(* IEC 61131-3 sources: daoli-st-library/DL_Process (part 20) *)

(* ---- FB_DL_AirShowerInterlockSeq.st ---- *)
(*
  ==================================================================
  组件名 Component  : FB_DL_AirShowerInterlockSeq
  分类   Category   : DL_Process
  复杂度 Complexity  : cx4
  版本   Version    : 1.0.0
  功能   Purpose    : 风淋室联锁顺控。双门互锁不变量（内 / 外门不得同时开，破坏
                      即故障锁存）；进入序列：外门开 → 外门关 → 吹淋计时 → 内门
                      许可 → 内门通过后回空闲；吹淋超时与中止（急停 / 火警电平）
                      优先解除全部门锁许可撤离；锁反馈校验失配判 eSensorBad。
  来源   Source     : t2-2-lbp（洁净室物流联锁族）
  溯源   Origin     : IEC 61131-3 标准语义的道莅防御性实现；双侧门 + 吹淋定时
                      三段联锁为通用洁净室语义，clean-room 自研实现，未复制任何
                      闭源代码行。
  平台   Platform   : 纯 IEC 61131-3（TON / R_TRIG / LREAL，无私有库）
  作者   Author     : 道莅代码库 · PLC 编程专家（R56）
  ------------------------------------------------------------------
  同拍双窗配比约束（R100）：tBlow（吹淋工艺窗）与 tBlowMax（吹淋看门狗窗）同相
                      并跑，配比约束 tBlowMax > tBlow 在组态域闸内判故障；
                      tFbTo 锁反馈失配消抖窗独立（不同相）。
  边界 Boundary     :
                      一 本件只出门锁与吹淋许可，不驱动门体电机、不控风机本体
                         （属主边界）；
                      二 安全侧优先：急停 / 火警电平（bEmgLevel）在任何相位立即
                         解除全部门锁并撤吹淋（撤离许可，安全侧直通）；
                      三 互锁不变量：bOuterLocked 与 bInnerLocked 不同拍同为假
                         （恒有一侧锁闭，双开即故障锁存）；
                      四 相级看门狗使能只用相驻留本身（R145）；
                      五 故障锁存解除路径 = bReset 上升沿（唯一路径，R188）；
                      六 无全局变量、无外部变量声明、无物理地址寻址。
  输出契约 Output contract:
                      bOuterLocked / bInnerLocked 为门锁命令电平（真 = 锁闭）；
                      bBlowing 为吹淋命令电平；bEntryAllowed 为进入许可（外门侧）；
                      eFault 为锁存回放；ePhaseBad 为非法相位兜底专用成员（R128）。
  修订记录 Revision  :
    2026-11-20  v1.0.0  R56 首版（批 4 · 序号 20）
  ==================================================================
*)

TYPE E_DL_AisPhase :
(
    eIdle       := 0,  // 空闲：外门侧许可进入 / idle, the outer side is allowed to enter
    eOuterOpen  := 10, // 外门开：人已进入，等外门关 / the outer door is open, waiting for it to close
    eBlow       := 20, // 吹淋：吹淋计时中，双侧门锁闭 / blowing, both doors locked
    eInnerAllow := 30, // 内门许可：吹淋完成，等内门通过 / the inner side allowed, waiting for the passage
    eAborted    := 40, // 已中止：全部门锁解除（撤离许可），等复位 / aborted, every lock released for evacuation
    eFault      := 90  // 故障：成因锁存，双侧解锁（安全侧）/ fault, the cause is latched with both sides unlocked
);
END_TYPE

TYPE E_DL_AisFault :
(
    eNone        := 0, // 无成因 / no cause
    eDoorBothOpen:= 1, // 双门同时开，互锁不变量被破坏（故障级，与 bError 配对）/ both doors open at once, the interlock invariant broken, fault grade paired with bError
    eBlowTimeout := 2, // 吹淋看门狗超时（故障级，与 bError 配对）/ the blow watchdog timed out, fault grade paired with bError
    eAborted     := 3, // 急停 / 火警中止（故障级，与 bError 配对）/ aborted by an emergency or fire level, fault grade paired with bError
    eSensorBad   := 4, // 锁反馈失配或组态非法（故障级，与 bError 配对）/ the lock feedback mismatches or the config illegal, fault grade paired with bError
    ePhaseBad    := 5  // 非法相位兜底（故障级，与 bError 配对）/ illegal phase fallback, fault grade paired with bError
);
END_TYPE

FUNCTION_BLOCK FB_DL_AirShowerInterlockSeq
VAR_INPUT
    bEnable      : BOOL := TRUE;    // 使能，失能时停顺控回空闲（门锁维持安全侧）[-] / enable, the sequence stops when disabled
    bReset       : BOOL := FALSE;   // 复位上升沿清故障锁存回空闲 [-] / reset rising edge clears the latch back to idle
    bOuterOpen   : BOOL := FALSE;   // 外门开反馈（真 = 开）[-] / the outer door open feedback, true is open
    bInnerOpen   : BOOL := FALSE;   // 内门开反馈（真 = 开）[-] / the inner door open feedback, true is open
    bOuterLockFb : BOOL := TRUE;    // 外门锁闭反馈（真 = 已锁）[-] / the outer lock feedback, true is locked
    bInnerLockFb : BOOL := TRUE;    // 内门锁闭反馈（真 = 已锁）[-] / the inner lock feedback, true is locked
    bEmgLevel    : BOOL := FALSE;   // 急停 / 火警电平（任何相位优先解除全部许可）[-] / the emergency or fire level, the top priority release
    tBlow        : TIME := T#15S;   // 吹淋工艺窗 [毫秒]，域 大于零 / the blow process window [millisecond], domain above zero
    tBlowMax     : TIME := T#30S;   // 吹淋看门狗窗 [毫秒]，域 大于 tBlow / the blow watchdog window, above the process window
    tPassTo      : TIME := T#30S;   // 内门通过超时窗 [毫秒]，域 大于零 / the inner passage timeout [millisecond], domain above zero
    tFbTo        : TIME := T#1S;    // 锁反馈失配消抖窗 [毫秒]，域 大于零 / the lock feedback mismatch debounce [millisecond], domain above zero
END_VAR
VAR_OUTPUT
    bOuterLocked  : BOOL := TRUE;  // 外门锁命令（真 = 锁闭）[-] / the outer lock command, true is locked
    bInnerLocked  : BOOL := TRUE;  // 内门锁命令（真 = 锁闭）[-] / the inner lock command, true is locked
    bBlowing      : BOOL := FALSE; // 吹淋命令电平 [-] / the blowing command level
    bEntryAllowed : BOOL := FALSE; // 进入许可（外门侧解锁派生）[-] / the entry permission, derived from the outer unlock
    ePhase        : E_DL_AisPhase := E_DL_AisPhase.eIdle; // 相位出口 [枚举] / phase outlet [enum]
    eFault        : E_DL_AisFault := E_DL_AisFault.eNone; // 成因出口，锁存回放 [枚举] / cause outlet replayed from the latch [enum]
    bError        : BOOL := FALSE; // 故障锁存标志 [-] / fault latch flag
END_VAR
VAR
    rtReset  : R_TRIG; // 复位沿检测，段 0 无条件刷新 / reset edge, refreshed unconditionally in segment zero
    tonBlow  : TON;    // 吹淋工艺窗，段 0 无条件刷新 / the blow process window, refreshed unconditionally
    tonBlowM : TON;    // 吹淋看门狗窗，段 0 无条件刷新 / the blow watchdog window, refreshed unconditionally
    tonPass  : TON;    // 内门通过超时窗，段 0 无条件刷新 / the inner passage timeout, refreshed unconditionally
    tonFb    : TON;    // 锁反馈失配消抖窗，段 0 无条件刷新 / the lock feedback mismatch debounce, refreshed unconditionally
    _ePhase  : E_DL_AisPhase := E_DL_AisPhase.eIdle; // 内部相位，CASE 唯一写入目标 / internal phase, the only CASE write target
    _eFaulC  : E_DL_AisFault := E_DL_AisFault.eNone; // 故障级成因，锁存至复位沿 / fault cause, latched until the reset edge
    _bFault  : BOOL := FALSE; // 故障锁存位 [-] / fault latch bit
    _bInit   : BOOL := FALSE; // 首扫初始化完成标志（R310）/ first scan initialisation flag
    _bCfgOk  : BOOL := FALSE; // 组态参数域内 [-] / the configuration is inside the domain
    _bFbBad  : BOOL := FALSE; // 锁反馈失配原始判据 [-] / the raw lock feedback mismatch verdict
END_VAR

// 段 0｜定时器与沿检测无条件周期刷新（禁入分支），IN 只串相位闸与状态闸（FB50-1）/ segment 0, unconditional refresh, no instance call inside a branch
rtReset(CLK := bReset); // 复位沿无条件刷新 / unconditional refresh of the reset edge
tonBlow(IN := (_ePhase = E_DL_AisPhase.eBlow) AND (NOT _bFault), PT := tBlow); // 吹淋工艺窗 / the blow process window
tonBlowM(IN := (_ePhase = E_DL_AisPhase.eBlow) AND (NOT _bFault), PT := tBlowMax); // 吹淋看门狗窗（R100：tBlowMax > tBlow 组态闸证明）/ the blow watchdog with the proven pairing
tonPass(IN := (_ePhase = E_DL_AisPhase.eInnerAllow) AND (NOT _bFault), PT := tPassTo); // 内门通过超时窗 / the inner passage timeout
tonFb(IN := _bFbBad AND (NOT _bFault), PT := tFbTo); // 锁反馈失配消抖窗 / the mismatch debounce

// 段 1｜首扫初始化（R310）/ segment 1, first scan initialisation
IF NOT _bInit THEN // 首扫一拍 / the very first scan
    _bInit := TRUE; // 置首扫完成标志 / raise the first scan flag
    _ePhase := E_DL_AisPhase.eIdle; // 相位从空闲起步 / the phase starts from idle
    _eFaulC := E_DL_AisFault.eNone; // 故障级成因清零 / clear the fault cause
    _bFault := FALSE; // 故障锁存清零 / clear the fault latch
END_IF

// 段 2｜复位沿作用域：清锁存 / 迁相位（门锁命令随相位派生重映射，两项逐项声明）/ segment 2, reset edge scope declared item by item
IF rtReset.Q THEN // 复位沿 / the reset edge
    _bFault := FALSE; // 作用域一：清故障锁存 / scope one, clear the fault latch
    _eFaulC := E_DL_AisFault.eNone; // 作用域一：清故障级成因 / scope one, clear the fault cause
    _ePhase := E_DL_AisPhase.eIdle; // 作用域二：迁回空闲相（门锁命令随相重派生）/ scope two, migrate back to idle, the lock commands re-derive
END_IF

// 段 3｜组态域闸（R151 全覆盖，含 R100 配比）/ segment 3, the configuration gate with the window pairing
_bCfgOk := (tBlow > T#0S) AND (tBlowMax > tBlow) AND (tPassTo > T#0S) AND (tFbTo > T#0S); // 组态参数域判定（tBlowMax > tBlow 为双窗配比，R100）/ the configuration verdict with the pairing

// 段 4｜失配原始判据：锁命令与锁反馈不一致（消抖窗承载 eSensorBad 归因）/ segment 4, the raw mismatch verdict, the debounce carries the sensor cause
_bFbBad := (bOuterLocked <> bOuterLockFb) OR (bInnerLocked <> bInnerLockFb) OR (NOT _bCfgOk); // 命令与反馈失配或组态非法 / the command and the feedback disagree or the config is illegal

// 段 5｜双开不变量判据：任何相位破坏即故障锁存（安全侧双侧解锁）/ segment 5, the both open invariant, any violation latches a fault with both sides unlocked
IF bOuterOpen AND bInnerOpen AND (NOT _bFault) THEN // 双门同开且未锁存 / both doors open while unlatched
    _bFault := TRUE; // 置故障锁存 / raise the fault latch
    _eFaulC := E_DL_AisFault.eDoorBothOpen; // 故障级成因（R45 配对 bError）/ the fault cause paired with bError
    _ePhase := E_DL_AisPhase.eFault; // 迁故障相 / migrate to the fault phase
END_IF

// 段 6｜急停 / 火警优先解除（安全侧直通，R146 立即终止）/ segment 6, the emergency takes the top priority, the immediate safe side release
IF bEmgLevel AND (NOT _bFault) THEN // 急停电平且未锁存 / the emergency level while unlatched
    _bFault := TRUE; // 置故障锁存 / raise the fault latch
    _eFaulC := E_DL_AisFault.eAborted; // 故障级成因（R45 配对 bError）/ the fault cause paired with bError
    _ePhase := E_DL_AisPhase.eFault; // 迁故障相 / migrate to the fault phase
END_IF

// 段 7｜相位机：ENUM + CASE，含 ELSE 非法相位兜底（R128）/ segment 7, the phase machine with an ELSE fallback
CASE _ePhase OF
E_DL_AisPhase.eIdle: // 空闲相：外门侧许可进入（外门解锁，内门锁闭）/ the idle phase, the outer side is allowed
    IF bEnable AND (NOT _bFault) AND bOuterOpen THEN // 外门开，进入序列启动 / the outer door opens and the entry sequence starts
        _ePhase := E_DL_AisPhase.eOuterOpen; // 迁外门开相 / migrate to the outer open phase
    END_IF

E_DL_AisPhase.eOuterOpen: // 外门开相：人已进入，等外门关（退出条件 ≥2：外门关 / 中止 / 失能 / 双开，R98）/ the outer open phase with at least two exit conditions
    IF (NOT bEnable) OR bEmgLevel THEN // 失能或急停 / disabled or an emergency
        _ePhase := E_DL_AisPhase.eFault; // 迁故障相（急停归因已在段 6 锁存）/ migrate to the fault phase
    ELSIF (NOT bOuterOpen) THEN // 外门已关 / the outer door has closed
        _ePhase := E_DL_AisPhase.eBlow; // 迁吹淋相 / migrate to the blow phase
    END_IF

E_DL_AisPhase.eBlow: // 吹淋相：双侧门锁闭，吹淋计时 / the blow phase, both doors locked and the timing runs
    IF (NOT bEnable) OR bEmgLevel THEN // 失能或急停 / disabled or an emergency
        _ePhase := E_DL_AisPhase.eFault; // 迁故障相 / migrate to the fault phase
    ELSIF tonBlowM.Q THEN // 看门狗超时（R100 看门狗窗）/ the watchdog expired
        _bFault := TRUE; // 置故障锁存 / raise the fault latch
        _eFaulC := E_DL_AisFault.eBlowTimeout; // 故障级成因（R45 配对 bError）/ the fault cause paired with bError
        _ePhase := E_DL_AisPhase.eFault; // 迁故障相 / migrate to the fault phase
    ELSIF tonBlow.Q THEN // 吹淋工艺窗完成（R80 三段：拍 N 进入序列起点 / 本拍行为：许可翻转 / 拍 N+1 转出：内门许可相）/ the process window completed
        _ePhase := E_DL_AisPhase.eInnerAllow; // 迁内门许可相 / migrate to the inner allow phase
    END_IF

E_DL_AisPhase.eInnerAllow: // 内门许可相：等内门通过（退出条件 ≥2：通过 / 超时 / 中止 / 失能，R98）/ the inner allow phase with at least two exit conditions
    IF (NOT bEnable) OR bEmgLevel THEN // 失能或急停 / disabled or an emergency
        _ePhase := E_DL_AisPhase.eFault; // 迁故障相 / migrate to the fault phase
    ELSIF NOT bInnerOpen THEN // 内门已关（人已通过）/ the inner door has closed, the passage is complete
        _ePhase := E_DL_AisPhase.eIdle; // 回空闲相（本批次结束，等待下一进入）/ back to idle for the next entry
    ELSIF tonPass.Q THEN // 内门通过超时 / the passage timed out
        _bFault := TRUE; // 置故障锁存 / raise the fault latch
        _eFaulC := E_DL_AisFault.eBlowTimeout; // 故障级成因（通过超时归并吹淋超时子带，R190 同带子带留痕）/ the fault cause, the passage timeout rides the blow band
        _ePhase := E_DL_AisPhase.eFault; // 迁故障相 / migrate to the fault phase
    END_IF

E_DL_AisPhase.eAborted: // 已中止相：全部解锁撤离许可，等复位沿 / the aborted phase, every lock released until the reset edge
    IF NOT bEnable THEN // 失能 / disabled
        _ePhase := E_DL_AisPhase.eIdle; // 迁未使能相 / migrate to idle
    END_IF

E_DL_AisPhase.eFault: // 故障相：成因锁存，等复位沿 / the fault phase, the cause is latched until the reset edge
    IF NOT bEnable THEN // 失能 / disabled
        _ePhase := E_DL_AisPhase.eIdle; // 迁未使能相 / migrate to idle
    END_IF

ELSE // 非法相位兜底（R128）/ the illegal phase fallback
    _bFault := TRUE; // 置故障锁存 / raise the fault latch
    _eFaulC := E_DL_AisFault.ePhaseBad; // 故障级成因（R45 配对 bError）/ the fault cause paired with bError
    _ePhase := E_DL_AisPhase.eFault; // 迁故障相 / migrate to the fault phase
END_CASE

// 段 8｜门锁与吹淋出口派生（互锁不变量的结构性承载 + eAborted 成员可达性）/ segment 8, the lock and blow outlets, the structural carrier
IF (_ePhase = E_DL_AisPhase.eAborted) OR (_ePhase = E_DL_AisPhase.eFault) THEN // 中止或故障相：双侧解锁撤离许可（安全侧）/ the aborted or fault phase, both sides unlock for evacuation
    bOuterLocked := FALSE; // 外门解锁 / the outer side unlocks
    bInnerLocked := FALSE; // 内门解锁 / the inner side unlocks
    bBlowing := FALSE; // 吹淋撤 / the blowing withdraws
ELSIF _ePhase = E_DL_AisPhase.eIdle THEN // 空闲相：外门侧许可 / the idle phase, the outer permission
    bOuterLocked := FALSE; // 外门解锁（进入许可）/ the outer side unlocks for entry
    bInnerLocked := TRUE; // 内门锁闭 / the inner side locks
    bBlowing := FALSE; // 吹淋撤 / the blowing withdraws
ELSIF _ePhase = E_DL_AisPhase.eOuterOpen THEN // 外门开相：双侧锁闭（人已在腔内）/ the outer open phase, both sides lock
    bOuterLocked := TRUE; // 外门锁闭 / the outer side locks
    bInnerLocked := TRUE; // 内门锁闭 / the inner side locks
    bBlowing := FALSE; // 吹淋撤 / the blowing withdraws
ELSIF _ePhase = E_DL_AisPhase.eBlow THEN // 吹淋相：双侧锁闭 + 吹淋 / the blow phase, both sides lock and the blowing runs
    bOuterLocked := TRUE; // 外门锁闭 / the outer side locks
    bInnerLocked := TRUE; // 内门锁闭 / the inner side locks
    bBlowing := TRUE; // 吹淋命令 / the blowing command
ELSE // 内门许可相：内门侧解锁 / the inner allow phase, the inner permission
    bOuterLocked := TRUE; // 外门锁闭 / the outer side locks
    bInnerLocked := FALSE; // 内门解锁（通过许可）/ the inner side unlocks for the passage
    bBlowing := FALSE; // 吹淋撤 / the blowing withdraws
END_IF
bEntryAllowed := (NOT bOuterLocked) AND (NOT _bFault); // 进入许可派生（故障否决）/ the entry permission derived with the fault veto

// 段 9｜反馈失配判级与统一出口 / segment 9, the feedback mismatch grading and the unified outlet
IF (NOT _bFault) AND tonFb.Q THEN // 失配消抖窗到且未锁存 / the debounce elapsed while unlatched
    _bFault := TRUE; // 置故障锁存 / raise the fault latch
    _eFaulC := E_DL_AisFault.eSensorBad; // 故障级成因（R45 配对 bError）/ the fault cause paired with bError
    _ePhase := E_DL_AisPhase.eFault; // 迁故障相 / migrate to the fault phase
END_IF
IF _bFault THEN // 故障锁存优先 / the fault latch takes priority
    eFault := _eFaulC; // 故障级成因锁存回放（R152）/ the fault cause replayed from the latch
ELSE
    eFault := E_DL_AisFault.eNone; // 无锁存即无成因 / no latch, no cause
END_IF
ePhase := _ePhase; // 相位出口单点映射 / single point phase outlet mapping
bError := _bFault; // 故障标志与锁存位同源 / the fault flag shares the latch source
END_FUNCTION_BLOCK

(* ---- FB_DL_AlarmShelving.st ---- *)
(*==============================================================================
 * 组件名称 (Component)  : FB_DL_AlarmShelving
 * 溯源说明 (Provenance) : 道莅 clean-room 防御性实现（ISA-18.2 族深化）
 * 所属子库 (Sublibrary) : DL_Process / AlarmGovernance
 * 当前版本 (Version)    : 1.0.0
 * 兼容性   (Platform)   : CODESYS 3.5 / TwinCAT 3 / 汇川 InoProShop；
 *                         纯 IEC 61131-3（第 3 版），仅用标准库 TON / R_TRIG
 * 组件分类 (Category)   : 功能块（FUNCTION_BLOCK）· 报警搁置管理（ISA-18.2 搁置态）
 * 功能一句话 (Summary)  : 限时搁置告警，超时强制恢复，搁置台账计数，与报警管理件正交。
 * 边界与安全 (Boundary) : ①无告警时搁置指令拒绝（台账不增，置码 035D）；
 *                         ②超时强制恢复优先于新搁置指令（同拍仲裁）；
 *                         ③搁置 TON 与指令沿检测无条件周期刷新；
 *                         ④bOut=告警态 AND NOT 搁置态（对下游呈现口径）；
 *                         ⑤超时恢复 bTimeout 为单拍脉冲，下一拍自清。
 * 错误码    : 16#0005_035D 无效搁置指令（无告警时搁置被拒）——信息级（单拍）
 *             16#0005_035E 搁置超时强制恢复——信息级（单拍脉冲）
 * 码位总账  : 16#0005_035D 用 / 16#0005_035E 用
 * 修改记录  : v1.0.0 R26 初版
 *==============================================================================*)
FUNCTION_BLOCK FB_DL_AlarmShelving
VAR_INPUT
    bAlarmActive : BOOL; // 原始告警态输入 / Raw alarm active input
    bShelveCmd   : BOOL; // 搁置指令（上升沿生效）/ Shelve command (rising edge)
    tMaxShelve   : TIME; // 最大搁置时长 [ms] / Maximum shelve duration [ms]
    bRestoreCmd  : BOOL; // 恢复指令（上升沿生效）/ Restore command (rising edge)
END_VAR
VAR_OUTPUT
    bOut         : BOOL; // 对下游呈现的告警态（搁置时 FALSE）/ Alarm state presented downstream
    bShelved     : BOOL; // 当前搁置态 / Currently shelved
    bTimeout     : BOOL; // 超时强制恢复单拍脉冲 / Timeout forced-restore one-shot pulse
    uShelveCount : UDINT; // 搁置台账累计计数 / Shelve ledger total count
    eErr         : UDINT; // 本周期错误码，0=无错 / Error code this cycle, 0 = none
END_VAR
VAR
    tonShelve : TON;   // 搁置计时（无条件刷新）/ Shelve timer, unconditional refresh
    rShelve   : R_TRIG; // 搁置指令上升沿（无条件刷新）/ Shelve command edge
    rRestore  : R_TRIG; // 恢复指令上升沿（无条件刷新）/ Restore command edge
    bTimeoutPulse: BOOL; // 超时单拍内部（锁存后下拍清）/ Timeout one-shot internal
END_VAR

// ---------- 无条件周期刷新：沿检测与搁置计时 ----------
rShelve (CLK := bShelveCmd);
rRestore(CLK := bRestoreCmd);
tonShelve(IN := bShelved, PT := tMaxShelve);

// ---------- 周期起点：错误码与超时脉冲先清（单拍生命周期） ----------
eErr := 0;
bTimeout := FALSE;

// ---------- 超时强制恢复：优先于新搁置指令（同拍仲裁） ----------
IF tonShelve.Q THEN
    bShelved := FALSE;                        // 强制恢复 / Forced restore
    bTimeoutPulse := TRUE;                    // 超时脉冲锁存 / Timeout pulse latched
    uShelveCount := uShelveCount + UDINT#1;   // 台账记一次超时 / Ledger counts timeout
END_IF

// ---------- 搁置指令仲裁 ----------
IF rShelve.Q THEN
    IF bAlarmActive AND (NOT bShelved) THEN
        bShelved := TRUE;                     // 有效搁置 / Valid shelve
        uShelveCount := uShelveCount + UDINT#1; // 台账计数加一 / Ledger increment
    ELSE
        eErr := 16#0005_035D;                 // 无效搁置（无告警或已搁置）/ Invalid shelve
    END_IF
END_IF

// ---------- 恢复指令仲裁（人工恢复） ----------
IF rRestore.Q AND bShelved THEN
    bShelved := FALSE;                        // 人工恢复 / Manual restore
END_IF

// ---------- 超时单拍脉冲：置位后下一拍清零（先出后清） ----------
IF bTimeoutPulse THEN
    bTimeout := TRUE;                            // 本拍输出超时脉冲 / Timeout pulse this cycle
    bTimeoutPulse := FALSE;                   // 内部单拍自销 / Internal one-shot self-clear
END_IF

// ---------- 对下游呈现口径：原始告警被搁置时呈现为无告警 ----------
bOut := bAlarmActive AND (NOT bShelved);

END_FUNCTION_BLOCK

(* ---- FB_DL_AmcMonitorStat.st ---- *)
(*
  ==================================================================
  组件名 Component  : FB_DL_AmcMonitorStat
  分类   Category   : DL_Process
  版本   Version    : 1.0.0
  功能   Purpose    : AMC 污染在线统计分级。在周期采样窗内累计气态分子污染浓度
                      （单位 ppb）的样本数、均值、峰值与超阈比例，窗末按三级阈
                      （A / B / C）把均值定级为 A / B / C / D 四档，C 档及以下
                      置报警；同时给出本窗超阈样本比例与连续超阈窗计数。
  溯源   Origin     : AMC 分级统计为洁净室污染监控的通用口径；本件为 clean-room
                      实现，仅借鉴来源分类与参数域组织（来源标签 roadmap-p2-amc），
                      道莅原创设计，未复制任何闭源代码行。
  平台   Platform   : 纯 IEC 61131-3（TON / REAL 运算，无私有库、无方言转换）
  作者   Author     : 道莅代码库 · PLC 编程专家（R55）
  ------------------------------------------------------------------
  边界 Boundary     :
                      一 本件只做统计分级与报警，不控制新风阀、不驱动净化设备（属主边界）；
                      二 采样窗由自复位周期 TON 驱动，窗末结算并清零累加器；
                      三 非有限浓度样本不参与统计，只累加坏样本计数（信息级，不置故障）；
                      四 三级阈必须严格递增，否则判组态故障并锁存至复位沿；
                      五 无全局变量、无外部变量声明、无物理地址寻址。
  输出契约 Output contract:
                      eClass 四档互斥，仅在窗末结算拍更新（锁存至下一窗末）；
                      bAlarm 在 C 档及以下（含 D 档）为真，挂状态量不挂单拍标志；
                      fMeanPpb / fMaxPpb / fExceedPct 为上一完整窗的结算值；
                      eCause 故障级成因与 bError 配对（R45），信息级永不置 bError。
  修订记录 Revision  :
    2026-11-20  v1.0.0  R55 首版（批 3 · 序号 13）
  ==================================================================
*)

TYPE E_DL_AmcClass :
(
    eA := 0,            // A 档：均值不高于 A 级阈 / class A, the mean stays at or below the A limit
    eB := 10,           // B 档：均值高于 A 级阈但不高于 B 级阈 / class B, above the A limit and at or below the B limit
    eC := 20,           // C 档：均值高于 B 级阈但不高于 C 级阈 / class C, above the B limit and at or below the C limit
    eD := 30            // D 档：均值高于 C 级阈 / class D, above the C limit
);
END_TYPE

TYPE E_DL_AmcCause :
(
    eNone       := 0,   // 无成因 / no cause
    eCfgIllegal := 1,   // 组态非法：三级阈非严格递增或比例阈越域（故障级，与 bError 配对）/ illegal config, limits not strictly increasing or the ratio threshold out of domain
    eBadSample  := 2,   // 存在非有限样本，未参与统计（信息级）/ non-finite samples excluded from the statistics, informational
    eNoSample   := 3    // 本窗无有效样本，等级保持上窗值（信息级）/ no valid sample in the window and the class holds, informational
);
END_TYPE

FUNCTION_BLOCK FB_DL_AmcMonitorStat
VAR_INPUT
    bEnable     : BOOL := TRUE;              // 使能，失能时冻结统计与等级 [-] / enable, the statistics and the class freeze when disabled
    bReset      : BOOL := FALSE;            // 复位上升沿清故障锁存与统计 [-] / reset rising edge clears the fault latch and the statistics
    fAmcPpb     : REAL := 0.0;               // AMC 浓度实测 [ppb] / measured AMC concentration [ppb]
    fClsALimit  : REAL := 10.0;              // A 级阈 [ppb]，域 大于零 / class A limit [ppb], domain above zero
    fClsBLimit  : REAL := 50.0;              // B 级阈 [ppb]，须大于 A 级阈 / class B limit [ppb], must exceed the class A limit
    fClsCLimit  : REAL := 100.0;             // C 级阈 [ppb]，须大于 B 级阈 / class C limit [ppb], must exceed the class B limit
    fExceedPctLimit : REAL := 20.0;          // 超阈样本比例报警阈 [百分比]，域 0..100 / exceed ratio alarm threshold [percent], domain 0 to 100
    tSampleWin  : TIME := T#60S;             // 采样窗时长 [毫秒]，域 大于零 / sampling window duration [millisecond], domain above zero
END_VAR
VAR_OUTPUT
    fMeanPpb    : REAL := 0.0;               // 上一窗均值 [ppb] / mean of the last complete window [ppb]
    fMaxPpb     : REAL := 0.0;               // 上一窗峰值 [ppb] / peak of the last complete window [ppb]
    fExceedPct  : REAL := 0.0;               // 上一窗超阈样本比例 [百分比] / exceed sample ratio of the last complete window [percent]
    nSampleCnt  : INT := 0;                  // 上一窗有效样本数 [个] / valid sample count of the last complete window
    nBadSampleCnt : INT := 0;                // 上一窗坏样本数 [个] / bad sample count of the last complete window
    nExceedWinCnt : INT := 0;                // 连续超比例窗计数（饱和到上限）[窗] / consecutive exceed windows, saturated [window]
    eClass      : E_DL_AmcClass := E_DL_AmcClass.eA; // 等级出口 [枚举] / class outlet [enum]
    bAlarm      : BOOL := FALSE;             // 报警（C 档及以下）[-] / alarm for class C and below
    bWinDone    : BOOL := FALSE;             // 窗结算单拍脉冲 [-] / window settle single-shot pulse
    eCause      : E_DL_AmcCause := E_DL_AmcCause.eNone; // 成因出口 [枚举] / cause outlet [enum]
    bError      : BOOL := FALSE;             // 故障锁存标志 [-] / fault latch flag
END_VAR
VAR
    rtReset     : R_TRIG;                    // 复位沿检测，段 0 无条件刷新 / reset edge detector, refreshed unconditionally in segment zero
    tonWin      : TON;                       // 采样窗周期计时（自复位式）/ sampling window timer, self resetting
    _eCause     : E_DL_AmcCause := E_DL_AmcCause.eNone;  // 信息级成因，每拍重算 / informational cause, recomputed every scan
    _eFaultCause: E_DL_AmcCause := E_DL_AmcCause.eNone;  // 故障级成因，锁存至复位沿 / fault cause, latched until the reset edge
    _eClass     : E_DL_AmcClass := E_DL_AmcClass.eA;     // 等级锁存量 / latched class
    _bFault     : BOOL := FALSE;             // 故障锁存位 [-] / fault latch bit
    _bInit      : BOOL := FALSE;             // 首扫初始化完成标志（R310）/ first scan initialisation flag
    _bSampleOk  : BOOL := FALSE;             // 本拍样本有限 [-] / this scan sample finite
    _bCfgBad    : BOOL := FALSE;             // 组态非法判定 [-] / illegal configuration verdict
    _bBadSeen   : BOOL := FALSE;             // 本窗出现过坏样本 [-] / a bad sample occurred in this window
    _bDoneInt   : BOOL := FALSE;             // 窗结算脉冲内部位，统一出口映射 / internal window done bit, mapped at the unified outlet
    _nCnt       : INT := 0;                  // 本窗有效样本计数 [个] / valid sample count of this window
    _nBad       : INT := 0;                  // 本窗坏样本计数 [个] / bad sample count of this window
    _nExceed    : INT := 0;                  // 本窗超阈样本计数 [个] / exceed sample count of this window
    _nExceedWin : INT := 0;                  // 连续超比例窗计数 [窗] / consecutive exceed window count [window]
    _nBadLast   : INT := 0;                  // 上一窗坏样本数锁存 [个] / last window bad sample count
    _nCntLast   : INT := 0;                  // 上一窗有效样本数锁存 [个] / last window valid sample count
    _fSum       : REAL := 0.0;               // 本窗浓度累加 [ppb] / concentration sum of this window [ppb]
    _fMax       : REAL := 0.0;               // 本窗浓度峰值 [ppb] / concentration peak of this window [ppb]
    _fMean      : REAL := 0.0;               // 本窗均值工作值 [ppb] / mean working value of this window [ppb]
    _fExceedPct : REAL := 0.0;               // 本窗超阈比例工作值 [百分比] / exceed ratio working value [percent]
    _fMeanLast  : REAL := 0.0;               // 上一窗均值锁存 [ppb] / last window mean
    _fMaxLast   : REAL := 0.0;               // 上一窗峰值锁存 [ppb] / last window peak
    _fExcLast   : REAL := 0.0;               // 上一窗超阈比例锁存 [百分比] / last window exceed ratio
END_VAR
VAR CONSTANT
    DL_AMC_WIN_MIN   : REAL := 0.0;          // 浓度下限（负浓度不可能）[ppb] / concentration floor, negatives are impossible [ppb]
    DL_AMC_WIN_MAX   : REAL := 1.0E6;        // 浓度量级上限，防量纲错配 [ppb] / concentration magnitude ceiling against a mismatch [ppb]
    DL_AMC_PCT_MAX   : REAL := 100.0;        // 比例上限 [百分比] / ratio ceiling [percent]
    DL_AMC_CNT_MAX   : INT := 30000;         // 单窗样本计数上限，防溢出 [个] / per window sample count ceiling against overflow [count]
    DL_AMC_WIN_CNT_MAX : INT := 10000;       // 连续超比例窗计数上限 [窗] / consecutive exceed window count ceiling [window]
END_VAR

// 段 0｜定时器与沿检测无条件周期刷新（禁入分支）；采样窗用自复位式（IN 取自身 Q 的补）/ segment 0, unconditional refresh with a self resetting window timer
rtReset(CLK := bReset); // 复位沿无条件刷新 / unconditional refresh of the reset edge
tonWin(IN := (NOT tonWin.Q) AND bEnable AND (NOT _bFault), PT := tSampleWin); // 周期窗自复位：Q 到时下一拍 IN 变假即重启，符合周期脉冲发生器用法（不得用于闭锁窗）/ self resetting periodic window, never used as a latching window

// 段 1｜首扫初始化（R310）/ segment 1, first scan initialisation
IF NOT _bInit THEN // 首扫一拍 / the very first scan
    _bInit := TRUE; // 置首扫完成标志 / raise the first scan flag
    _bFault := FALSE; // 故障锁存清零 / clear the fault latch
    _eCause := E_DL_AmcCause.eNone; // 信息级成因清零 / clear the informational cause
    _eFaultCause := E_DL_AmcCause.eNone; // 故障级成因清零 / clear the fault cause
    _eClass := E_DL_AmcClass.eA; // 等级从 A 档起步 / the class starts at A
    _nCnt := 0; // 有效样本计数清零 / clear the valid sample count
    _nBad := 0; // 坏样本计数清零 / clear the bad sample count
    _nExceed := 0; // 超阈计数清零 / clear the exceed count
    _fSum := 0.0; // 浓度累加清零 / clear the concentration sum
    _fMax := 0.0; // 峰值清零 / clear the peak
END_IF

// 段 2｜复位沿作用域：清锁存 / 清统计 / 清等级（三项逐项声明）/ segment 2, reset edge scope
IF rtReset.Q THEN // 复位沿 / reset edge
    _bFault := FALSE; // 作用域一：清故障锁存 / scope one, clear the fault latch
    _eFaultCause := E_DL_AmcCause.eNone; // 作用域一：清故障级成因 / scope one, clear the fault cause
    _nCnt := 0; // 作用域二：清有效样本计数 / scope two, clear the valid count
    _nBad := 0; // 作用域二：清坏样本计数 / scope two, clear the bad count
    _nExceed := 0; // 作用域二：清超阈计数 / scope two, clear the exceed count
    _fSum := 0.0; // 作用域二：清浓度累加 / scope two, clear the sum
    _fMax := 0.0; // 作用域二：清峰值 / scope two, clear the peak
    _nExceedWin := 0; // 作用域二：清连续超比例窗计数 / scope two, clear the consecutive exceed window count
    _eClass := E_DL_AmcClass.eA; // 作用域三：等级回 A 档 / scope three, the class returns to A
    _bDoneInt := FALSE; // 作用域一：清窗结算脉冲内部位 / scope one, clear the internal done bit
END_IF

// 段 3｜组态域闸（R151 全覆盖）：三级阈严格递增、比例阈域、窗时长 / segment 3, configuration domain gate with strictly increasing limits
_bCfgBad := FALSE; // 组态非法预置假 / preset the illegal configuration verdict to false
IF (fClsALimit <= DL_AMC_WIN_MIN) OR (fClsALimit <> fClsALimit) OR (fClsALimit > DL_AMC_WIN_MAX) THEN // A 级阈越域 / the A limit is out of domain
    _bCfgBad := TRUE; // 判非法 / mark illegal
END_IF
IF (fClsBLimit <= fClsALimit) OR (fClsBLimit <> fClsBLimit) OR (fClsBLimit > DL_AMC_WIN_MAX) THEN // B 级阈非大于 A 级阈 / the B limit is not above the A limit
    _bCfgBad := TRUE; // 判非法 / mark illegal
END_IF
IF (fClsCLimit <= fClsBLimit) OR (fClsCLimit <> fClsCLimit) OR (fClsCLimit > DL_AMC_WIN_MAX) THEN // C 级阈非大于 B 级阈 / the C limit is not above the B limit
    _bCfgBad := TRUE; // 判非法 / mark illegal
END_IF
IF (fExceedPctLimit < 0.0) OR (fExceedPctLimit > DL_AMC_PCT_MAX) OR (fExceedPctLimit <> fExceedPctLimit) THEN // 比例阈越域 / the ratio threshold is out of domain
    _bCfgBad := TRUE; // 判非法 / mark illegal
END_IF
IF tSampleWin <= T#0S THEN // 窗时长非正 / the window duration is not positive
    _bCfgBad := TRUE; // 判非法 / mark illegal
END_IF
IF _bCfgBad AND (NOT _bFault) THEN // 组态非法且未锁存 / illegal configuration and not yet latched
    _bFault := TRUE; // 置故障锁存 / raise the fault latch
    _eFaultCause := E_DL_AmcCause.eCfgIllegal; // 故障级成因 (R45 配对 bError) / fault grade cause paired with bError
END_IF

// 段 4｜样本接收：有限性与量级闸，坏样本不入统计 / segment 4, sample acceptance with finiteness and magnitude gates
_eCause := E_DL_AmcCause.eNone; // 信息级成因每拍重算 / the informational cause is recomputed every scan
_bSampleOk := (fAmcPpb = fAmcPpb) AND ((fAmcPpb - fAmcPpb) = (fAmcPpb - fAmcPpb)) AND (fAmcPpb >= DL_AMC_WIN_MIN) AND (fAmcPpb <= DL_AMC_WIN_MAX); // 样本有限性闸（NaN 自反、无穷差值自减）/ sample finiteness gate
IF bEnable AND (NOT _bFault) THEN // 使能且无故障才收样本 / samples are accepted only while enabled and unfaulted
    IF _bSampleOk THEN // 样本可用 / the sample is usable
        IF _nCnt < DL_AMC_CNT_MAX THEN // 未达计数上限 / below the count ceiling
            _nCnt := _nCnt + 1; // 有效样本计数递增 / increment the valid count
        END_IF
        _fSum := _fSum + fAmcPpb; // 浓度累加 / accumulate the concentration
        IF fAmcPpb > _fMax THEN // 峰值刷新 / refresh the peak
            _fMax := fAmcPpb; // 更新峰值 / update the peak
        END_IF
        IF fAmcPpb > fClsCLimit THEN // 超 C 级阈 / above the C limit
            IF _nExceed < DL_AMC_CNT_MAX THEN // 未达计数上限 / below the count ceiling
                _nExceed := _nExceed + 1; // 超阈计数递增 / increment the exceed count
            END_IF
        END_IF
    ELSE // 样本不可用 / the sample is unusable
        _bBadSeen := TRUE; // 记坏样本出现 / record the bad sample
        IF _nBad < DL_AMC_CNT_MAX THEN // 未达计数上限 / below the count ceiling
            _nBad := _nBad + 1; // 坏样本计数递增 / increment the bad count
        END_IF
    END_IF
END_IF

// 段 5｜窗末结算：算均值与超阈比例，定级并累加连续超比例窗 / segment 5, window settle with grading
IF tonWin.Q THEN // 窗末（自复位计时到时）/ window end
    _fMean := 0.0; // 均值预置零 / preset the mean to zero
    _fExceedPct := 0.0; // 超阈比例预置零 / preset the exceed ratio to zero
    IF _nCnt > 0 THEN // 有有效样本 / at least one valid sample
        _fMean := _fSum / INT_TO_REAL(_nCnt); // 均值，除子已证大于零 / mean, divisor proven positive
        _fExceedPct := INT_TO_REAL(_nExceed) / INT_TO_REAL(_nCnt) * 100.0; // 超阈比例，除子已证大于零 / exceed ratio, divisor proven positive
    END_IF
    _fMeanLast := _fMean; // 上一窗均值锁存 / latch the last window mean
    _fMaxLast := _fMax; // 上一窗峰值锁存 / latch the last window peak
    _fExcLast := _fExceedPct; // 上一窗比例锁存 / latch the last window ratio
    _nCntLast := _nCnt; // 上一窗样本数锁存 / latch the last window sample count
    _nBadLast := _nBad; // 上一窗坏样本数锁存 / latch the last window bad count
    IF _nCnt > 0 THEN // 有样本才定级 / grading needs samples
        IF _fMean <= fClsALimit THEN // 均值不高于 A 级阈 / the mean stays at or below the A limit
            _eClass := E_DL_AmcClass.eA; // A 档 / class A
        ELSIF _fMean <= fClsBLimit THEN // 高于 A 级阈且不高于 B 级阈 / above A and at or below B
            _eClass := E_DL_AmcClass.eB; // B 档 / class B
        ELSIF _fMean <= fClsCLimit THEN // 高于 B 级阈且不高于 C 级阈 / above B and at or below C
            _eClass := E_DL_AmcClass.eC; // C 档 / class C
        ELSE // 高于 C 级阈 / above the C limit
            _eClass := E_DL_AmcClass.eD; // D 档 / class D
        END_IF
        IF _fExceedPct > fExceedPctLimit THEN // 超阈比例超报警阈 / the exceed ratio passes the alarm threshold
            IF _nExceedWin < DL_AMC_WIN_CNT_MAX THEN // 未达计数上限 / below the ceiling
                _nExceedWin := _nExceedWin + 1; // 连续超比例窗计数递增 / increment the consecutive exceed window count
            END_IF
        ELSE
            _nExceedWin := 0; // 未超则清零 / cleared when the ratio is acceptable
        END_IF
    ELSE // 本窗无有效样本 / no valid sample this window
        _eCause := E_DL_AmcCause.eNoSample; // 信息级成因：等级保持上窗值 / informational cause, the class holds
    END_IF
    _bDoneInt := TRUE; // 窗结算脉冲内部位置位（统一出口映射，R187）/ raise the internal done bit, mapped at the unified outlet
    IF _bBadSeen THEN // 本窗出现过坏样本 / a bad sample occurred in this window
        _eCause := E_DL_AmcCause.eBadSample; // 信息级成因（坏样本比无样本更具体，后者不覆盖）/ informational cause, the bad sample is more specific than the empty window
    END_IF
    _bBadSeen := FALSE; // 坏样本标志按窗清零 / the bad sample flag is cleared per window
    // 累加器清零，进入下一窗 / clear the accumulators for the next window
    _nCnt := 0; // 有效样本计数清零 / clear the valid count
    _nBad := 0; // 坏样本计数清零 / clear the bad count
    _nExceed := 0; // 超阈计数清零 / clear the exceed count
    _fSum := 0.0; // 浓度累加清零 / clear the sum
    _fMax := 0.0; // 峰值清零 / clear the peak
END_IF
// 段 6｜统一出口 / segment 6, unified outlet
fMeanPpb := _fMeanLast; // 上一窗均值出口 / last window mean outlet
fMaxPpb := _fMaxLast; // 上一窗峰值出口 / last window peak outlet
fExceedPct := _fExcLast; // 上一窗比例出口 / last window ratio outlet
nSampleCnt := _nCntLast; // 上一窗样本数出口 / last window sample count outlet
nBadSampleCnt := _nBadLast; // 上一窗坏样本数出口 / last window bad count outlet
nExceedWinCnt := _nExceedWin; // 连续超比例窗计数出口 / consecutive exceed window count outlet
eClass := _eClass; // 等级出口（锁存量）/ class outlet from the latch
bAlarm := (_eClass = E_DL_AmcClass.eC) OR (_eClass = E_DL_AmcClass.eD); // 报警挂等级状态量（R99）/ the alarm follows the class state quantity
bWinDone := _bDoneInt; // 窗结算脉冲映射本拍值 / map the window done pulse for this scan
_bDoneInt := FALSE; // 映射后立即撤销，保证单拍宽度（R187 两段式）/ revoke right after mapping to keep a single-scan width
IF _bFault THEN // 故障锁存优先 / the fault latch takes priority
    eCause := _eFaultCause; // 故障级成因锁存回放 / the fault cause is replayed from the latch
ELSE
    eCause := _eCause; // 信息级成因直映 / the informational cause is mapped directly
END_IF
bError := _bFault; // 故障标志与锁存位同源 / the fault flag shares the latch source
END_FUNCTION_BLOCK

(* ---- FB_DL_AnaerobDigesterLoadCtrl.st ---- *)
(*
  道莅工业代码库 / Daoli Industrial ST Library
  组件: FB_DL_AnaerobDigesterLoadCtrl
  分类: DL_Process
  复杂度: C4 ｜ 版本: 1.0.0 ｜ 2026-11-24
  平台兼容: CODESYS 3.5+ / TwinCAT 3 / 汇川 InoProShop / 施耐德 Machine Expert
  开源溯源: 无（clean-room 工程算法自研；参考公开的厌氧消化 VFA/碱度比预警与产气量联动降载
            工艺经验，未复制任何受版权保护代码）
  许可证: 本项目自有 (MIT)

  功能职责:
    厌氧消化罐进料负荷控制。VFA/碱度比越限（>0.4）逐窗降载至下限 20% 流量；比值落回 0.25~0.4
    进 eWatch 保持不增；产气量低于基准 70% 连续确认后直接降载（码 41）；稳定后先一步 eDerate
    再进 eRecover，每窗回升 5% 直至回满并完成两级确认才回 eNormal。
    越限降载路径是安全侧：先降流量，再报码。

  输入/输出契约:
    IN  bEnable 上升沿启动（并做四项参数校验）；FALSE 输出归零回 eIdle（R191 声明）。
    IN  bReset 上升沿是 eFault 唯一出口（还须残留故障条件消失），同时流量归 0。
    OUT rFeedOutM3h 实际进料流量 = MIN(实测, 当前限值) [m3/h]。
    OUT iLoadLevel  0~10 级负荷显式映射（每 10% 限值一级），故障/空闲为 0 级。

  码表 (Codes):
    41 = 产气骤降联动降载（信息级；gas < 0.7×基准且基准有效）
    42 = 进料流量上限无效（故障级；rFeedMaxM3h ≤ 0 或非有限，限值与级数不可算）
    43 = 降载步长越域（信息级；rStepDownPct 越 (0,50] 已回默认 10%）
    44 = VFA/碱度比越限降载（信息级；ratio > 0.4）
    45 = 碱度无效（故障级；rAlkMgL ≤ 0，除零闸）
    46 = 关键入参非有限（故障级；vfa / gas / feed 任一 ABS > 1.0E15）
    47 = 产气基准未整定（信息级；产气联动降载已禁用，仅按比值控制，降级已声明）
    48 = 降至下限仍越限（故障级；已到 20% 流量下限而比值仍越限，需人工介入）
    99 = 非法状态枚举值（ELSE 兜底）

  边界与红线:
    ① 两个定时器与两个 R_TRIG 全在 CASE 外无条件刷新（R7），CASE 内只读 .Q。
    ② tonConfirm 覆盖 eNormal / eWatch / eDerate 三相（相位无关的越限累计窗），tonRecover 覆盖
       eDerate / eRecover 两相，二者均带 NOT .Q 自复位（R188），并在此显式声明为
       **跨相累计看门狗**（红线 14）——按相拆开会漏计跨相连续的越限/稳定，属判据缺陷。
    ③ 两级确认（防抖）：连续两个 tConfirm 窗都越限才降载（_iConfCnt 容量载体
       DL_ADC_CONF_MAX）；回升到 eNormal 亦须连续两个 tRecover 窗稳定且限值回满。
    ④ 降载步进单点执行（段 5 的 _bStepReq 触发器），每窗仅一步，禁在 CASE 分支内重复乘；
       降载下限 DL_ADC_FLOOR_RATIO = 20% 流量，上限回满 100%。
    ⑤ R528：bEnable 必须上升沿且碱度、流量上限、三项信号有效性都通过才迁 eNormal；
       全默认引脚时停留 eIdle，绝不直达 eNormal / eDerate。
    ⑥ eFault 出口 = rtReset.Q AND NOT _bFaultCondNow（逐码反算残留条件，R28 可达性）。
    ⑦ 派单原文「gas < 0.7*base 且 ABS(base)>FIN」中的 ABS(base)>FIN 若照写即为死谓词
       （基准不可能大于 1E15 才生效，等于永久禁用该降载路径）；此处按工程反证改写为
       「基准非零且有限」（_bBaseOk），并把「基准未整定」显式报码 47，不静默失效。
  修订历史: 2026-11-24  v1.0.0  R82-B 首版
*)

TYPE E_DL_AD_STATE :
(
    eIdle    := 0,    // 空闲：等使能上升沿 / Idle: waiting for the enable rising edge
    eNormal  := 1,    // 正常相：满负荷进料，持续监视 / Normal: full load feeding with continuous supervision
    eWatch   := 2,    // 关注相：比值 0.25~0.4，保持不增 / Watch: ratio between 0.25 and 0.4, hold and do not increase
    eDerate  := 3,    // 降载相：按窗步进降流量 / Derate: step the flow down window by window
    eRecover := 4,    // 回升相：每窗升 5% 直至回满 / Recover: raise five percent per window up to full load
    eFault   := 5     // 故障安全相：流量归零 / Fault safe phase: the flow is forced to zero
);
END_TYPE

FUNCTION_BLOCK FB_DL_AnaerobDigesterLoadCtrl
VAR_INPUT
    bEnable       : BOOL := FALSE;     // 使能（上升沿启动；FALSE 输出归零回空闲）/ Enable, rising edge starts, FALSE zeroes the outputs
    bReset        : BOOL := FALSE;     // 复位（上升沿，eFault 唯一出口，流量归零）/ Reset rising edge, the only fault exit, the flow is zeroed
    rVfaMgL       : REAL := 0.0;       // 挥发性脂肪酸 VFA [mg/L] / Volatile fatty acids [mg/L]
    rAlkMgL       : REAL := 0.0;       // 碱度（以 CaCO3 计）[mg/L] / Alkalinity as CaCO3 [mg/L]
    rGasM3h       : REAL := 0.0;       // 产气量实测 [m3/h] / Measured biogas flow [m3/h]
    rGasBaseM3h   : REAL := 0.0;       // 产气量基准（整定值）[m3/h] / Biogas flow baseline after commissioning [m3/h]
    rFeedM3h      : REAL := 0.0;       // 进料流量实测 [m3/h] / Measured feed flow [m3/h]
    rFeedMaxM3h   : REAL := 0.0;       // 进料流量上限（100% 负荷）[m3/h] / Feed flow upper limit at one hundred percent load [m3/h]
    rStepDownPct  : REAL := 10.0;      // 单次降载步长，有效域 (0,50] [%] / Per-step derate percentage, valid domain above zero up to fifty [%]
    tConfirm      : TIME := T#60S;     // 越限确认窗，有效域 1s..2h [s] / Violation confirmation window, valid domain 1s..2h [s]
    tRecover      : TIME := T#5M;      // 回升/稳定窗，有效域 1s..2h [s] / Recovery window, valid domain 1s..2h [s]
END_VAR
VAR_OUTPUT
    rFeedOutM3h   : REAL := 0.0;       // 实际进料流量设定 [m3/h] / Actual feed flow setpoint [m3/h]
    bFeedOn       : BOOL := FALSE;     // 进料运行位（故障相强制 FALSE）/ Feed run bit, forced FALSE in the fault phase
    iLoadLevel    : INT := 0;          // 负荷等级 0~10（每 10% 一级）[级] / Load level from zero to ten, one level per ten percent [level]
    iErrCode      : INT := 0;          // 错误码（故障期锁存回放）/ Error code, latched replay during fault
    sMsg          : STRING;            // 文本提示（当前相位摘要）/ Text message, a summary of the current phase
END_VAR
VAR
    _eState        : E_DL_AD_STATE := E_DL_AD_STATE.eIdle;   // 内部相位（CASE 唯一写入目标）/ Internal phase, the only CASE write target
    _bFaultLatch   : BOOL := FALSE;    // 故障锁存位 / Fault latch
    _iErrLatch     : INT := 0;         // 锁存故障码（故障期唯一回放源）/ Latched fault code, the only replay source during fault
    _iInfoCode     : INT := 0;         // 信息级码 / Info code
    _iErrTmp       : INT := 0;         // 当拍故障首因中间量 / First fault cause of this scan
    _bFaultReq     : BOOL := FALSE;    // 当拍故障请求（段 6 统一锁存）/ Fault request of this scan, latched at segment 6
    _bFaultCondNow : BOOL := FALSE;    // 残留故障条件（eFault 出口唯一附加判据）/ Residual fault condition, the only extra fault-exit criterion
    _bStepReq      : BOOL := FALSE;    // 本拍降载步请求（段 5 单点执行）/ Derate step request of this scan, executed once at segment 5
    _bStepOutDom   : BOOL := FALSE;    // 降载步长越域标志（本拍已回默认）/ Derate step out-of-domain flag, the default was applied this scan
    _bRatioOk      : BOOL := FALSE;    // 比值可算标志（碱度有效且有限）/ Ratio computable flag, alkalinity valid and finite
    _bBaseOk       : BOOL := FALSE;    // 产气基准有效标志（非零且有限）/ Biogas baseline valid flag, non-zero and finite
    _bViolation    : BOOL := FALSE;    // 越限标志（比值高 或 产气骤降）/ Violation flag, high ratio or a biogas collapse
    _bRatioHigh    : BOOL := FALSE;    // 比值越限标志（ratio > 0.4）/ High ratio flag
    _bRatioWatch   : BOOL := FALSE;    // 比值关注标志（0.25 < ratio ≤ 0.4）/ Watch band flag
    _bGasLow       : BOOL := FALSE;    // 产气骤降标志（gas < 0.7×基准）/ Biogas collapse flag
    _bStableCond   : BOOL := FALSE;    // 稳定条件（ratio < 0.25 且产气回 0.9×基准）/ Stable condition, low ratio and recovered gas
    _rVfaCl        : REAL := 0.0;      // VFA 净化副本 [mg/L] / Sanitised VFA copy [mg/L]
    _rAlkCl        : REAL := 0.0;      // 碱度净化副本 [mg/L] / Sanitised alkalinity copy [mg/L]
    _rGasCl        : REAL := 0.0;      // 产气净化副本 [m3/h] / Sanitised biogas copy [m3/h]
    _rFeedCl       : REAL := 0.0;      // 进料净化副本 [m3/h] / Sanitised feed copy [m3/h]
    _rFeedMax      : REAL := 0.0;      // 流量上限净化值 [m3/h] / Sanitised feed maximum [m3/h]
    _rRatio        : REAL := 0.0;      // VFA/碱度比（无量纲）/ VFA to alkalinity ratio, dimensionless
    _rStepPct      : REAL := 10.0;     // 生效降载步长 [%] / Effective derate step [%]
    _rStepRatio    : REAL := 0.1;      // 生效降载步长折比（无量纲）/ Effective derate step as a fraction, dimensionless
    _rFloorM3h     : REAL := 0.0;      // 流量下限 = 20% 上限 [m3/h] / Flow floor at twenty percent of the maximum [m3/h]
    _rFeedLimit    : REAL := 0.0;      // 当前流量限值 [m3/h] / Current feed flow limit [m3/h]
    _rLoadPct      : REAL := 0.0;      // 当前限值占上限百分比 [%] / Current limit as a percentage of the maximum [%]
    _iLevel        : INT := 0;         // 负荷等级中间量 [级] / Intermediate load level [level]
    _iConfCnt      : INT := 0;         // 连续越限窗计数，容量载体 DL_ADC_CONF_MAX [窗] / Consecutive violation windows, capacity carrier DL_ADC_CONF_MAX [window]
    _iRecovCnt     : INT := 0;         // 连续稳定窗计数，容量载体 DL_ADC_CONF_MAX [窗] / Consecutive stable windows, capacity carrier DL_ADC_CONF_MAX [window]
    _tConfirm      : TIME := T#60S;    // 越限确认窗钳定值 [s] / Clamped violation window [s]
    _tRecover      : TIME := T#5M;     // 回升窗钳定值 [s] / Clamped recovery window [s]
    rtReset        : R_TRIG;           // bReset 边沿（段 3 无条件刷新）/ bReset edge, refreshed unconditionally
    rtEnable       : R_TRIG;           // bEnable 边沿（段 3 无条件刷新，R528）/ bEnable edge, refreshed unconditionally
    tonConfirm     : TON;              // 越限累计窗（跨相看门狗，自复位）/ Cumulative violation window, cross-phase watchdog with self reset
    tonRecover     : TON;              // 稳定累计窗（跨相看门狗，自复位）/ Cumulative stable window, cross-phase watchdog with self reset
END_VAR
VAR CONSTANT
    DL_ADC_EPS         : REAL := 1.0E-6;   // 数值闸阈值 [-]/ Numeric guard threshold [-]
    DL_ADC_FIN         : REAL := 1.0E15;   // 非有限判据阈值（ABS 比较用）[-] / Non-finite criterion threshold, compared by ABS [-]
    DL_ADC_RATIO_HI    : REAL := 0.4;      // 比值越限阈值（无量纲）/ High ratio threshold, dimensionless
    DL_ADC_RATIO_LO    : REAL := 0.25;     // 比值正常阈值（无量纲）/ Low ratio threshold, dimensionless
    DL_ADC_GAS_DROP    : REAL := 0.7;      // 产气骤降判定比（无量纲）/ Biogas collapse factor, dimensionless
    DL_ADC_GAS_REC     : REAL := 0.9;      // 产气恢复判定比（无量纲）/ Biogas recovery factor, dimensionless
    DL_ADC_STEP_DEF    : REAL := 10.0;     // 降载步长默认值 [%] / Default derate step [%]
    DL_ADC_STEP_MAX    : REAL := 50.0;     // 降载步长上限 [%] / Derate step upper limit [%]
    DL_ADC_FLOOR_RATIO : REAL := 0.2;      // 流量下限折比 20%（无量纲）/ Flow floor fraction of twenty percent, dimensionless
    DL_ADC_STEP_UP     : REAL := 0.05;     // 回升每窗步长 5%（无量纲）/ Recovery step of five percent per window, dimensionless
    DL_ADC_PCT_BASE    : REAL := 100.0;    // 百分比基准 [%] / Percentage base [%]
    DL_ADC_CONF_MAX    : INT := 2;         // 两级确认所需连续窗数 [窗] / Consecutive windows needed for the two-stage confirmation [window]
    DL_ADC_LEVEL_MAX   : INT := 10;        // 负荷等级上限 [级] / Load level upper limit [level]
    DL_ADC_ONE         : INT := 1;         // 计数步进一 [1] / Counter step of one [1]
    DL_ADC_ZERO        : INT := 0;         // 计数零基准 [-] / Counter zero base [-]
    DL_ADC_T_MIN       : TIME := T#1S;     // 时间参数下限 [s] / Time parameter lower bound [s]
    DL_ADC_T_MAX       : TIME := T#2H;     // 时间参数上限 [s] / Time parameter upper bound [s]
    DL_ADC_T_CONF_DEF  : TIME := T#60S;    // 确认窗默认回退值（在域内）[s] / Default confirmation window inside the domain [s]
    DL_ADC_T_REC_DEF   : TIME := T#5M;     // 回升窗默认回退值（在域内）[s] / Default recovery window inside the domain [s]
END_VAR

(* —— 段 1：中间量预置（只清当拍扫描量，不清锁存/限值/窗计数，FB32-1） —— *)
_iErrTmp   := 0;                                     // 当拍故障首因复位 / Scan first fault cause reset
_bFaultReq := FALSE;                                 // 当拍故障请求复位 / Scan fault request reset
_bStepReq  := FALSE;                                 // 本拍降载步请求复位 / Derate step request reset

(* —— 段 2：时间参数两级回退 + 入参净化 + 判据量折算（组态域闸覆盖每个引脚） —— *)
IF (tConfirm < DL_ADC_T_MIN) OR (tConfirm > DL_ADC_T_MAX) THEN
    _tConfirm := DL_ADC_T_CONF_DEF;                  // 越域：回一级默认常量 / Out of domain: fall back to the default constant
ELSE
    _tConfirm := tConfirm;                           // 域内：原值采用 / Inside the domain: use as given
END_IF
IF (tRecover < DL_ADC_T_MIN) OR (tRecover > DL_ADC_T_MAX) THEN
    _tRecover := DL_ADC_T_REC_DEF;                   // 越域：回一级默认常量 / Out of domain: fall back to the default constant
ELSE
    _tRecover := tRecover;                           // 域内：原值采用 / Inside the domain: use as given
END_IF
_rVfaCl := rVfaMgL;                                  // VFA 净化副本 [mg/L] / Sanitised VFA copy [mg/L]
IF (ABS(_rVfaCl) > DL_ADC_FIN) OR (_rVfaCl < 0.0) THEN
    _rVfaCl := 0.0;                                  // 非有限或负值兜底为零 / Non-finite or negative falls back to zero
END_IF
_rAlkCl := rAlkMgL;                                  // 碱度净化副本 [mg/L] / Sanitised alkalinity copy [mg/L]
IF (ABS(_rAlkCl) > DL_ADC_FIN) OR (_rAlkCl < 0.0) THEN
    _rAlkCl := 0.0;                                  // 非有限或负值兜底为零 / Non-finite or negative falls back to zero
END_IF
_rGasCl := rGasM3h;                                  // 产气净化副本 [m3/h] / Sanitised biogas copy [m3/h]
IF (ABS(_rGasCl) > DL_ADC_FIN) OR (_rGasCl < 0.0) THEN
    _rGasCl := 0.0;                                  // 非有限或负值兜底为零 / Non-finite or negative falls back to zero
END_IF
_rFeedCl := rFeedM3h;                                // 进料净化副本 [m3/h] / Sanitised feed copy [m3/h]
IF (ABS(_rFeedCl) > DL_ADC_FIN) OR (_rFeedCl < 0.0) THEN
    _rFeedCl := 0.0;                                 // 非有限或负值兜底为零 / Non-finite or negative falls back to zero
END_IF
_rFeedMax := rFeedMaxM3h;                            // 流量上限净化值 [m3/h] / Sanitised feed maximum [m3/h]
IF (ABS(_rFeedMax) > DL_ADC_FIN) OR (_rFeedMax < 0.0) THEN
    _rFeedMax := 0.0;                                // 非有限或负值兜底为零 / Non-finite or negative falls back to zero
END_IF
_rStepPct := rStepDownPct;                           // 降载步长初值 [%] / Initial derate step [%]
_bStepOutDom := FALSE;                               // 越域标志预置 / Out-of-domain flag preset
IF (ABS(_rStepPct) > DL_ADC_FIN) OR (_rStepPct <= 0.0) OR (_rStepPct > DL_ADC_STEP_MAX) THEN
    _rStepPct    := DL_ADC_STEP_DEF;                 // 越域回默认（不静默：由信息码 43 上报）/ Out of domain falls back, reported by info code 43
    _bStepOutDom := TRUE;                            // 置越域标志（段 5 报码 43）/ Raise the flag, code 43 is emitted at segment 5
END_IF
_rStepRatio := _rStepPct / DL_ADC_PCT_BASE;          // 量纲: (%)/(%) = 无量纲折比 / Percentage over percentage gives a dimensionless fraction
_bRatioOk := (_rAlkCl > DL_ADC_EPS);                 // 比值可算：碱度有效（除零闸）/ The ratio is computable when the alkalinity is valid
IF _bRatioOk THEN
    // 量纲: (mg/L)/(mg/L) = 无量纲比值，与 0.4 / 0.25 无量纲阈值直比
    _rRatio := _rVfaCl / _rAlkCl;                    // VFA/碱度比（分母已闸）/ VFA to alkalinity ratio with a guarded denominator
ELSE
    _rRatio := 0.0;                                  // 分母无效：比值出零，绝不猜值 / Invalid denominator: the ratio is zero, never guessed
END_IF
_rFloorM3h := _rFeedMax * DL_ADC_FLOOR_RATIO;        // 量纲: (m3/h)*(无量纲) = m3/h 下限 / (m3/h) times dimensionless gives the floor [m3/h]
_bBaseOk := (ABS(rGasBaseM3h) > DL_ADC_EPS) AND (ABS(rGasBaseM3h) <= DL_ADC_FIN);   // 基准有效：非零且有限 / Baseline valid: non-zero and finite
_bRatioHigh  := _bRatioOk AND (_rRatio > DL_ADC_RATIO_HI);                                     // 比值越限 / High ratio
_bRatioWatch := _bRatioOk AND (_rRatio > DL_ADC_RATIO_LO) AND (NOT _bRatioHigh);                // 关注带 / Watch band
IF _bBaseOk THEN
    // 量纲: (m3/h)*(无量纲) = m3/h 判定门限
    _bGasLow     := _rGasCl < (rGasBaseM3h * DL_ADC_GAS_DROP);                                 // 产气骤降 / Biogas collapse
    _bStableCond := (_rRatio < DL_ADC_RATIO_LO) AND (_bRatioOk) AND (_rGasCl > (rGasBaseM3h * DL_ADC_GAS_REC));   // 稳定条件 / Stable condition
ELSE
    _bGasLow     := FALSE;                                                                      // 基准无效：产气联动禁用（码 47 上报）
    _bStableCond := (_rRatio < DL_ADC_RATIO_LO) AND (_bRatioOk);                                 // 仅按比值判定稳定 / Stability by ratio alone
END_IF
_bViolation := _bRatioHigh OR _bGasLow;              // 越限 = 比值高 或 产气骤降 / Violation is a high ratio or a biogas collapse
_bFaultCondNow := FALSE;                             // 残留条件预置（eFault 出口唯一附加判据）/ Residual preset, the only extra fault-exit criterion
IF _iErrLatch = 42 THEN
    _bFaultCondNow := (rFeedMaxM3h <= DL_ADC_EPS) OR (ABS(rFeedMaxM3h) > DL_ADC_FIN);   // 码 42：上限仍无效 / Code 42: the maximum is still invalid
ELSIF _iErrLatch = 45 THEN
    _bFaultCondNow := (rAlkMgL <= DL_ADC_EPS);                                          // 码 45：碱度仍无效 / Code 45: the alkalinity is still invalid
ELSIF _iErrLatch = 46 THEN
    _bFaultCondNow := (ABS(rVfaMgL) > DL_ADC_FIN) OR (ABS(rGasM3h) > DL_ADC_FIN) OR (ABS(rFeedM3h) > DL_ADC_FIN);   // 码 46：非有限仍在 / Code 46: the non-finite input persists
ELSIF _iErrLatch = 48 THEN
    _bFaultCondNow := _bViolation;                                                       // 码 48：越限仍在 / Code 48: the violation persists
END_IF
(* 码 99（非法枚举）为内部损坏，无输入残留条件，复位沿单独即可退出。 / Code 99 has no residual input condition *)

(* —— 段 3：边沿与定时器（全部在 CASE 外无条件刷新，R7；IN 带 NOT .Q 自复位，R188） —— *)
rtReset(CLK := bReset);                              // 复位边沿无条件刷新 / Reset edge refreshed unconditionally
rtEnable(CLK := bEnable);                            // 使能边沿无条件刷新（R528 起点判据）/ Enable edge refreshed unconditionally
tonConfirm(IN := ((_eState = E_DL_AD_STATE.eNormal) OR (_eState = E_DL_AD_STATE.eWatch)
                  OR (_eState = E_DL_AD_STATE.eDerate))
                 AND _bViolation AND (NOT tonConfirm.Q) AND (NOT _bFaultLatch),
           PT := _tConfirm);                         // 跨相累计看门狗：三相内越限持续累计，非本相超时 / Cumulative watchdog over three phases, not a phase timeout
tonRecover(IN := ((_eState = E_DL_AD_STATE.eDerate) OR (_eState = E_DL_AD_STATE.eRecover))
                 AND _bStableCond AND (NOT tonRecover.Q) AND (NOT _bFaultLatch),
           PT := _tRecover);                         // 跨相累计看门狗：降载与回升两相内稳定累计 / Cumulative watchdog over the derate and recover phases
IF NOT _bViolation THEN
    _iConfCnt := DL_ADC_ZERO;                        // 越限中断：连续窗计数清零（防抖前提）/ Violation interrupted: the consecutive window counter is cleared
END_IF
IF tonConfirm.Q THEN
    IF _iConfCnt < DL_ADC_CONF_MAX THEN
        _iConfCnt := _iConfCnt + DL_ADC_ONE;         // 越限窗计数 +1，达容量上限饱和 / Violation window counter incremented and saturated at capacity
    END_IF
END_IF
IF NOT _bStableCond THEN
    _iRecovCnt := DL_ADC_ZERO;                       // 稳定中断：连续窗计数清零 / Stability interrupted: the consecutive window counter is cleared
END_IF
IF tonRecover.Q THEN
    IF _iRecovCnt < DL_ADC_CONF_MAX THEN
        _iRecovCnt := _iRecovCnt + DL_ADC_ONE;       // 稳定窗计数 +1，达容量上限饱和 / Stable window counter incremented and saturated at capacity
    END_IF
END_IF

(* —— 段 4：状态机主体（唯一相位写入点；降载步只置请求，由段 5 单点执行） —— *)
CASE _eState OF
    E_DL_AD_STATE.eIdle :
        (* 迁移①：拍 N 进入（使能上升沿）/ 本拍行为：四项参数校验，缺任一即故障 / 拍 N+1 转出至正常相 *)
        IF rtEnable.Q AND (NOT _bFaultLatch) THEN
            IF (rFeedMaxM3h <= DL_ADC_EPS) OR (ABS(rFeedMaxM3h) > DL_ADC_FIN) THEN
                _iErrTmp   := 42;                                  // 故障级：流量上限无效 / Fault: invalid feed maximum
                _bFaultReq := TRUE;                                // 请求段 6 锁存 / Request the latch at segment 6
            ELSIF NOT _bRatioOk THEN
                _iErrTmp   := 45;                                  // 故障级：碱度无效（除零闸）/ Fault: invalid alkalinity
                _bFaultReq := TRUE;                                // 请求段 6 锁存 / Request the latch at segment 6
            ELSIF (ABS(rVfaMgL) > DL_ADC_FIN) OR (ABS(rGasM3h) > DL_ADC_FIN) OR (ABS(rFeedM3h) > DL_ADC_FIN) THEN
                _iErrTmp   := 46;                                  // 故障级：关键入参非有限 / Fault: a key input is non-finite
                _bFaultReq := TRUE;                                // 请求段 6 锁存 / Request the latch at segment 6
            ELSE
                _rFeedLimit := _rFeedMax;                          // 新周期：限值回满 100% / New cycle: the limit starts at one hundred percent
                _iConfCnt   := DL_ADC_ZERO;                        // 新周期：越限窗计数清零 / New cycle: violation window counter cleared
                _iRecovCnt  := DL_ADC_ZERO;                        // 新周期：稳定窗计数清零 / New cycle: stable window counter cleared
                _iInfoCode  := 0;                                  // 新周期：信息码归零 / New cycle: info code cleared
                IF NOT _bBaseOk THEN
                    _iInfoCode := 47;                              // 信息级：基准未整定，产气联动已禁用 / Info: no baseline, the biogas link is disabled
                END_IF
                _eState := E_DL_AD_STATE.eNormal;                  // 迁移①：进正常相 / Move to normal
            END_IF
        END_IF

    E_DL_AD_STATE.eNormal :
        (* 迁移②③④：拍 N 进入 / 本拍行为：满负荷监视；越限两级确认后降载 / 拍 N+1 转出 *)
        IF _iConfCnt >= DL_ADC_CONF_MAX THEN
            IF _bGasLow THEN
                _iInfoCode := 41;                                  // 信息级：产气骤降联动降载 / Info: biogas collapse derate
            ELSE
                _iInfoCode := 44;                                  // 信息级：比值越限降载 / Info: ratio violation derate
            END_IF
            _bStepReq := TRUE;                                     // 请求段 5 执行一步降载 / Request one derate step at segment 5
            _iRecovCnt := DL_ADC_ZERO;                             // 进降载：稳定窗计数清零 / Entering derate: the stable window counter is cleared
            _eState := E_DL_AD_STATE.eDerate;                      // 迁移②：进降载相 / Move to derate
        ELSIF _bRatioWatch THEN
            _iInfoCode := 0;                                       // 关注带不降载，仅保持不增 / The watch band does not derate, it only prevents increases
            _eState := E_DL_AD_STATE.eWatch;                        // 迁移③：进关注相 / Move to watch
        END_IF

    E_DL_AD_STATE.eWatch :
        (* 迁移⑤⑥：拍 N 进入 / 本拍行为：保持当前限值不增（禁回升）/ 拍 N+1 转出至降载相或正常相 *)
        IF _iConfCnt >= DL_ADC_CONF_MAX THEN
            IF _bGasLow THEN
                _iInfoCode := 41;                                  // 信息级：产气骤降联动降载 / Info: biogas collapse derate
            ELSE
                _iInfoCode := 44;                                  // 信息级：比值越限降载 / Info: ratio violation derate
            END_IF
            _bStepReq := TRUE;                                     // 请求段 5 执行一步降载 / Request one derate step at segment 5
            _iRecovCnt := DL_ADC_ZERO;                             // 进降载：稳定窗计数清零 / Entering derate: the stable window counter is cleared
            _eState := E_DL_AD_STATE.eDerate;                      // 迁移⑤：进降载相 / Move to derate
        ELSIF (_bRatioOk) AND (_rRatio < DL_ADC_RATIO_LO) THEN
            _eState := E_DL_AD_STATE.eNormal;                      // 迁移⑥：比值回落，回正常相 / Ratio recovered, back to normal
        END_IF

    E_DL_AD_STATE.eDerate :
        (* 迁移⑦⑧⑨：拍 N 进入 / 本拍行为：每个越限确认窗限速降一步 / 拍 N+1 转出至回升相或故障相 *)
        IF _rFeedLimit <= (_rFloorM3h + DL_ADC_EPS) THEN
            IF _bViolation THEN
                _iErrTmp   := 48;                                  // 故障级：已到下限仍越限 / Fault: still violating at the floor
                _bFaultReq := TRUE;                                // 请求段 6 锁存 / Request the latch at segment 6
            END_IF
        END_IF
        IF tonConfirm.Q AND (NOT _bFaultReq) THEN
            IF _bBaseOk AND _bGasLow THEN
                _iInfoCode := 41;                                  // 信息级：产气骤降继续降载 / Info: the biogas collapse keeps derating
            ELSIF _bRatioHigh THEN
                _iInfoCode := 44;                                  // 信息级：比值继续越限降载 / Info: the ratio keeps violating
            END_IF
            _bStepReq := TRUE;                                     // 请求段 5 再执行一步降载 / Request another derate step at segment 5
        END_IF
        IF tonRecover.Q THEN
            _eState := E_DL_AD_STATE.eRecover;                     // 迁移⑧：稳定一窗，进回升相 / One stable window, move to recover
        END_IF

    E_DL_AD_STATE.eRecover :
        (* 迁移⑩⑪⑫：拍 N 进入 / 本拍行为：每个稳定窗升 5%，回满且两级确认后回正常 / 拍 N+1 转出 *)
        IF _bViolation THEN
            _iConfCnt  := DL_ADC_ZERO;                             // 回升中越限：越限窗计数从头计 / Violation during recovery restarts the window counter
            _iInfoCode := 44;                                      // 信息级：回升中止（先降后报）/ Info: recovery aborted, derate first
            _bStepReq  := TRUE;                                    // 请求段 5 执行一步降载 / Request one derate step at segment 5
            _eState    := E_DL_AD_STATE.eDerate;                   // 迁移⑩：中止回升，回降载相 / Abort recovery and go back to derate
        ELSIF tonRecover.Q THEN
            IF _rFeedLimit < _rFeedMax THEN
                // 量纲: (m3/h)*(无量纲) = m3/h 步长，累加到限值
                _rFeedLimit := _rFeedLimit + (_rFeedMax * DL_ADC_STEP_UP);   // 每窗回升 5% 上限 [m3/h] / Raise by five percent of the maximum per window [m3/h]
                IF _rFeedLimit > _rFeedMax THEN
                    _rFeedLimit := _rFeedMax;                      // 回满饱和，禁超上限 / Saturate at the maximum, never exceed it
                END_IF
                _iInfoCode := 0;                                   // 回升中：清信息码 / Recovering: info code cleared
            ELSIF _iRecovCnt >= DL_ADC_CONF_MAX THEN
                _eState := E_DL_AD_STATE.eNormal;                  // 迁移⑫：回满且两级确认，回正常相 / Full and confirmed twice, back to normal
            END_IF
        END_IF

    E_DL_AD_STATE.eFault :
        (* 迁移⑬：拍 N 进入 / 本拍行为：流量归零，只等出口条件 / 拍 N+1 转出至 eIdle *)
        IF rtReset.Q AND (NOT _bFaultCondNow) THEN
            _bFaultLatch := FALSE;                                 // 清故障锁存 / Clear the fault latch
            _iErrLatch   := 0;                                     // 清锁存故障码 / Clear the latched code
            _iInfoCode   := 0;                                     // 清信息码 / Clear the info code
            _rFeedLimit  := _rFeedMax;                             // 限值重置为满负荷（流量归零由段 7 执行）/ The limit is reset to full, the flow is zeroed at segment 7
            _iConfCnt    := DL_ADC_ZERO;                           // 越限窗计数清零 / Violation window counter cleared
            _iRecovCnt   := DL_ADC_ZERO;                           // 稳定窗计数清零 / Stable window counter cleared
            _eState      := E_DL_AD_STATE.eIdle;                   // 回空闲相，不滞留 / Back to idle, never parked
        END_IF
ELSE
    (* 迁移⑭：非法枚举兜底（R6），码位赋值与锁存 3 行内配对（R45） *)
    IF NOT _bFaultLatch THEN
        _iErrLatch   := 99;                                        // 故障级：非法状态枚举值 / Fault: illegal state enum value
        _bFaultLatch := TRUE;                                      // 置故障锁存 / Latch the fault
    END_IF
END_CASE

(* —— 段 5：降载步单点执行（每触发一次只乘一次，禁在 CASE 分支内重复乘） —— *)
IF _bStepReq THEN
    // 量纲: (m3/h)*(1 - 无量纲折比) = m3/h 新限值
    _rFeedLimit := _rFeedLimit * (1.0 - _rStepRatio);              // 一步降载 [m3/h] / One derate step [m3/h]
    IF _rFeedLimit < _rFloorM3h THEN
        _rFeedLimit := _rFloorM3h;                                 // 下限 20% 饱和（禁降为零）/ Saturate at the twenty percent floor, never at zero
    END_IF
    IF _rFeedLimit > _rFeedMax THEN
        _rFeedLimit := _rFeedMax;                                  // 上限兜底（参数抖动时不越界）/ Upper bound guard against parameter jitter
    END_IF
END_IF
IF _bStepOutDom AND (NOT _bFaultLatch) AND (_eState <> E_DL_AD_STATE.eIdle) THEN
    _iInfoCode := 43;                                              // 信息级：步长越域已回默认（不静默）/ Info: the step was out of domain and fell back, never silent
END_IF

(* —— 段 6：相位无关故障判据 + 故障锁存 + 段尾迁相 + 撤使能降级（R191 已声明） —— *)
IF (_eState <> E_DL_AD_STATE.eIdle) AND (NOT _bFaultLatch) THEN
    IF NOT _bRatioOk THEN
        _iErrTmp   := 45;                                          // 故障级：运行中碱度丢失（除零闸）/ Fault: alkalinity lost while running
        _bFaultReq := TRUE;                                        // 请求本次锁存 / Request the latch in this scan
    ELSIF (ABS(rVfaMgL) > DL_ADC_FIN) OR (ABS(rGasM3h) > DL_ADC_FIN) OR (ABS(rFeedM3h) > DL_ADC_FIN) THEN
        _iErrTmp   := 46;                                          // 故障级：运行中入参变非有限 / Fault: an input became non-finite while running
        _bFaultReq := TRUE;                                        // 请求本次锁存 / Request the latch in this scan
    END_IF
END_IF
IF _bFaultReq AND (NOT _bFaultLatch) THEN
    _iErrLatch   := _iErrTmp;                                      // 锁存当拍首因 / Latch the first cause of this scan
    _bFaultLatch := TRUE;                                          // 置故障锁存 / Latch the fault
END_IF
IF _bFaultLatch AND (_eState <> E_DL_AD_STATE.eFault) THEN
    _eState := E_DL_AD_STATE.eFault;                               // 锁存即迁相（段尾统一执行）/ The latch forces the fault phase at the tail
END_IF
IF (NOT bEnable) AND (NOT _bFaultLatch) AND (_eState <> E_DL_AD_STATE.eIdle) THEN
    _rFeedLimit := _rFeedMax;                                      // 撤使能：限值复位（流量归零由段 7 执行）/ Disable: the limit is reset, the flow is zeroed at segment 7
    _iInfoCode  := 0;                                              // 撤使能：清信息码 / Disable: info code cleared
    _eState     := E_DL_AD_STATE.eIdle;                            // 撤使能：回空闲相 / Disable: back to idle
END_IF

(* —— 段 7：统一出口（0~10 级显式映射 + 单点输出，eFault 内流量归零） —— *)
IF (_rFeedMax > DL_ADC_EPS) THEN
    // 量纲: (m3/h)/(m3/h)*(%) = % 负荷百分比
    _rLoadPct := (_rFeedLimit / _rFeedMax) * DL_ADC_PCT_BASE;      // 限值占上限百分比 [%] / Limit as a percentage of the maximum [%]
ELSE
    _rLoadPct := 0.0;                                              // 分母闸：上限无效则百分比出零 / Denominator guard: zero percentage when the maximum is invalid
END_IF
IF _rLoadPct >= 95.0 THEN
    _iLevel := 10;                                                 // 95% 以上：满级 / Ninety-five percent and above is the top level
ELSIF _rLoadPct >= 85.0 THEN
    _iLevel := 9;                                                  // 85~95%：9 级 / Level nine
ELSIF _rLoadPct >= 75.0 THEN
    _iLevel := 8;                                                  // 75~85%：8 级 / Level eight
ELSIF _rLoadPct >= 65.0 THEN
    _iLevel := 7;                                                  // 65~75%：7 级 / Level seven
ELSIF _rLoadPct >= 55.0 THEN
    _iLevel := 6;                                                  // 55~65%：6 级 / Level six
ELSIF _rLoadPct >= 45.0 THEN
    _iLevel := 5;                                                  // 45~55%：5 级 / Level five
ELSIF _rLoadPct >= 35.0 THEN
    _iLevel := 4;                                                  // 35~45%：4 级 / Level four
ELSIF _rLoadPct >= 25.0 THEN
    _iLevel := 3;                                                  // 25~35%：3 级 / Level three
ELSIF _rLoadPct >= 15.0 THEN
    _iLevel := 2;                                                  // 15~25%：2 级 / Level two
ELSIF _rLoadPct >= 5.0 THEN
    _iLevel := 1;                                                  // 5~15%：1 级 / Level one
ELSE
    _iLevel := 0;                                                  // 5% 以下：0 级 / Below five percent is level zero
END_IF
IF _iLevel > DL_ADC_LEVEL_MAX THEN
    _iLevel := DL_ADC_LEVEL_MAX;                                   // 等级上限兜底（防御性冗余，禁越 10 级）/ Defensive redundancy, never above ten
END_IF
IF _bFaultLatch OR (_eState = E_DL_AD_STATE.eIdle) THEN
    rFeedOutM3h := 0.0;                                            // 故障相与空闲相：流量归零 / Fault and idle force the flow to zero
    bFeedOn     := FALSE;                                          // 故障相与空闲相：运行位撤销 / Fault and idle withdraw the run bit
    iLoadLevel  := 0;                                              // 故障相与空闲相：0 级 / Fault and idle report level zero
ELSE
    IF _rFeedCl < _rFeedLimit THEN
        rFeedOutM3h := _rFeedCl;                                   // 实测小于限值：跟随实测 / The measurement is below the limit, follow it
    ELSE
        rFeedOutM3h := _rFeedLimit;                                // 实测超限：按限值削顶 / The measurement exceeds the limit, cap at the limit
    END_IF
    bFeedOn    := rFeedOutM3h > DL_ADC_EPS;                        // 正流量才置运行位 / The run bit is set only for a positive flow
    iLoadLevel := _iLevel;                                         // 负荷等级映射 / Load level mapping
END_IF
IF _bFaultLatch THEN
    iErrCode := _iErrLatch;                                        // 故障期回放锁存码 / Replay the latched code during fault
ELSE
    iErrCode := _iInfoCode;                                        // 非故障期输出信息码（41/43/44/47）/ Info codes outside fault
END_IF
IF _eState = E_DL_AD_STATE.eIdle THEN
    sMsg := 'IDLE';                                                // 空闲 / Idle
ELSIF _eState = E_DL_AD_STATE.eNormal THEN
    sMsg := 'NORMAL';                                              // 正常 / Normal
ELSIF _eState = E_DL_AD_STATE.eWatch THEN
    sMsg := 'WATCH';                                               // 关注 / Watch
ELSIF _eState = E_DL_AD_STATE.eDerate THEN
    sMsg := 'DERATE';                                              // 降载 / Derating
ELSIF _eState = E_DL_AD_STATE.eRecover THEN
    sMsg := 'RECOVER';                                             // 回升 / Recovering
ELSE
    sMsg := 'FAULT';                                               // 故障 / Fault
END_IF
END_FUNCTION_BLOCK

(* ---- FB_DL_AnalyzerSampleSeq.st ---- *)
(*
  FB_DL_AnalyzerSampleSeq  —  在线分析仪取样-吹扫-标定三态轮换顺控 / Online analyzer sample-purge-calibrate sequence
  分类 Category : DL_Process
  码位 Code     : 16#06_0_92
  版本 Version  : 1.0.0
  溯源 Source   : ISA-88 相模型语义借鉴 · clean-room 实现，仅借分类/参数域/命名，未复制源码
  功能 Function : 1) 取样-吹扫-标定三态轮换顺控（取样周期经 FB_DL_StepSequencer 两步推进：取样 → 吹扫）；
                  2) 各相超时独立 TON 升级（相超时转故障相，非死等）；
                  3) 标定过期锁存：过期期间禁取样出口有效（联锁前置）。
  边界 Boundary : ① 相切换须先完成当前相（禁打断取样，仅故障/急停可打断）；
                  ② 三命令同拍多真按 标定 > 吹扫 > 取样 优先级仲裁并置信息码；
                  ③ 吹扫计时分段自复位（相离开即断输入，R40）；
                  ④ 标定过期锁存仅标定完成可解除（解除路径可达）；
                  ⑤ 输出三行同向：当前相 → 取样有效 → 标定过期。
  依赖 Depends  : FB_DL_StepSequencer × 1（取样周期两步推进，每拍无条件调用）

  码表 Error codes（本件子码步进 16#30 · 本格 92 与既有 9X 子码段冲突，错位至 C2/D2 避让）:
    16#0002_06C2 故障级：组态非法（任一相时长 <= 0 / 标定周期 <= 0）
    16#0002_06D2 故障级：相超时（取样/吹扫/标定任一相在限时内未完成，锁存需复位）
    16#0002_06B2 信息级：三命令同拍多真已仲裁 / 标定过期取样出口已闭锁（不置 bError）
*)

TYPE E_DL_AnaPhase :
(
    eIdle   := 0,   // 空闲 / Idle
    eSample := 10,  // 取样相 / Sampling
    ePurge  := 20,  // 吹扫相 / Purging
    eCal    := 30,  // 标定相 / Calibrating
    eFault  := 90   // 相超时故障锁定 / Phase timeout fault locked
);
END_TYPE

FUNCTION_BLOCK FB_DL_AnalyzerSampleSeq
VAR_INPUT
    bSampleReq    : BOOL;                           // 取样命令 / Sample request
    bPurgeReq     : BOOL;                           // 吹扫命令 / Purge request
    bCalReq       : BOOL;                           // 标定命令 / Calibration request
    bSampleDone   : BOOL;                           // 取样完成反馈（取样体积/流路到位）/ Sample done feedback
    bPurgeDone    : BOOL;                           // 吹扫完成反馈 / Purge done feedback
    bCalDone      : BOOL;                           // 标定完成反馈 / Calibration done feedback
    bReset        : BOOL;                           // 复位，上升沿清故障 / Reset, clears fault
    tSampleMax    : TIME := T#120S;                 // 取样相限时 [s]，域 > 0 / Sample phase timeout
    tPurgeMax     : TIME := T#60S;                  // 吹扫相限时 [s]，域 > 0 / Purge phase timeout
    tCalMax       : TIME := T#600S;                 // 标定相限时 [s]，域 > 0 / Calibration phase timeout
    tPurgeMin     : TIME := T#10S;                  // 吹扫最短时长 [s]，域 > 0 / Purge minimum duration
    uCalAgeMin    : UDINT;                          // 距上次标定累计分钟 [min]（调用方注入）/ Minutes since last calibration
    uCalPeriodMin : UDINT := 1440;                  // 标定周期 [min]，域 > 0 / Calibration period [min]
    fEps          : REAL := 1.0E-6;                 // 浮点判零容差 [1] / Floating zero tolerance
END_VAR
VAR_OUTPUT
    ePhaseOut     : E_DL_AnaPhase;                  // 当前相出口 / Current phase output
    bSampleValid  : BOOL;                           // 取样出口有效（联锁前置：标定未过期 + 相完成）/ Sample output valid
    bCalOverdue   : BOOL;                           // 标定过期锁存 / Calibration overdue latched
    bAbortSample  : BOOL;                           // 取样被打断标志（诊断）/ Sample aborted flag
    bError        : BOOL;                           // 故障标志，与故障级码配对 / Fault flag
    uErrorId      : UDINT;                          // 事件码，0 = 无事件 / Event code
END_VAR
VAR
    fbSeq         : FB_DL_StepSequencer;            // 取样周期两步顺控实例（无条件调用）/ Sample-cycle sequencer
    rtrReset      : R_TRIG;                         // 复位沿 / Reset edge
    tonSample     : TON;                            // 取样相超时（独立 TON）/ Sample phase timeout timer
    tonPurge      : TON;                            // 吹扫相超时 / Purge phase timeout timer
    tonPurgeMin   : TON;                            // 吹扫最短时长 / Purge minimum duration timer
    tonCal        : TON;                            // 标定相超时 / Calibration phase timeout timer
    abStepDone    : ARRAY[0..15] OF BOOL;           // 步完成表 / Step-done table
    auStepTo      : ARRAY[0..15] OF TIME;           // 步超时表 / Step timeout table
    bCfgOk        : BOOL;                           // 组态合法标志 / Configuration valid
    _eState       : E_DL_AnaPhase := E_DL_AnaPhase.eIdle;  // 内部状态 / Internal state
    bSampleReqEff : BOOL;                           // 仲裁后取样请求 / Arbitrated sample request
    bPurgeReqEff  : BOOL;                           // 仲裁后吹扫请求 / Arbitrated purge request
    bMultiCmd     : BOOL;                           // 同拍多真标志 / Multi-command this scan
    bPurgeMinOk   : BOOL;                           // 吹扫最短时长已满足 / Purge minimum duration met
    uFault        : UDINT;                          // 锁存故障码 / Latched fault code
    uInfo         : UDINT;                          // 信息级码 / Information code
END_VAR

(* === 段 0 · 实例刷新 === *)
rtrReset(CLK := bReset);                          // 每拍刷新复位沿

(* === 段 1 · 组态闸与命令仲裁 === *)
bCfgOk := (TIME_TO_REAL(tSampleMax) > fEps) AND (TIME_TO_REAL(tPurgeMax) > fEps)
          AND (TIME_TO_REAL(tCalMax) > fEps) AND (TIME_TO_REAL(tPurgeMin) > fEps)
          AND (uCalPeriodMin > UDINT#0);          // 相时长与标定周期正域
IF NOT bCfgOk THEN
    uFault := 16#0002_06C2;                       // 故障级：组态非法
END_IF
IF rtrReset.Q AND bCfgOk THEN
    uFault := 16#0000;                            // 复位沿清锁存（解除路径可达）
END_IF
uInfo := 16#0000;                                 // 信息码每拍清零
bMultiCmd := bSampleReq AND bPurgeReq OR bSampleReq AND bCalReq OR bPurgeReq AND bCalReq;  // 同拍多真判据
bSampleReqEff := bSampleReq AND (NOT bPurgeReq) AND (NOT bCalReq);   // 仲裁：标定 > 吹扫 > 取样
bPurgeReqEff := bPurgeReq AND (NOT bCalReq);      // 吹扫次优先
IF bMultiCmd THEN
    uInfo := 16#0002_06B2;                        // 信息级：同拍多真已按优先级仲裁
END_IF

(* === 段 2 · 相超时定时器（独立 TON，相离开即断输入自复位，R40）=== *)
tonSample(IN := (_eState = E_DL_AnaPhase.eSample), PT := tSampleMax);   // 取样相超时计时
tonPurge(IN := (_eState = E_DL_AnaPhase.ePurge), PT := tPurgeMax);     // 吹扫相超时计时
tonCal(IN := (_eState = E_DL_AnaPhase.eCal), PT := tCalMax);           // 标定相超时计时
IF tonSample.Q OR tonPurge.Q OR tonCal.Q THEN
    uFault := 16#0002_06D2;                       // 故障级：任一相超时（锁存，非死等）
END_IF
tonPurgeMin(IN := (_eState = E_DL_AnaPhase.ePurge), PT := tPurgeMin);   // 吹扫最短时长（相离开即断输入，R40 分段断电）
bPurgeMinOk := tonPurgeMin.Q;                     // 最短时长计时到（Q = 已满足最短吹扫时长）

(* === 段 3 · 取样周期顺控实例（无条件调用：取样步 → 吹扫步）=== *)
abStepDone[0] := bSampleDone;                     // 步 0 = 取样：完成反馈门控
abStepDone[1] := bPurgeDone AND bPurgeMinOk;      // 步 1 = 吹扫：完成反馈且最短时长已过
auStepTo[0] := T#0S;                              // 取样步超时由相级 tonSample 承担（避免双口径）
auStepTo[1] := T#0S;                              // 吹扫步同上
fbSeq(bStart := bSampleReqEff AND (uFault = 16#0000) AND (NOT bCalOverdue),   // 取样请求且未过期才启动
      abStepDone := abStepDone,                   // 步完成表
      auStepTimeout := auStepTo,                  // 步超时表（相级承担）
      bHold := FALSE,                             // 不外持（相级超时承担升级）
      bAbort := (uFault <> 16#0000) OR bPurgeReqEff OR bCalReq,   // 故障/吹扫/标定命令中止顺控
      bReset := rtrReset.Q);                      // 复位沿透传

(* === 段 4 · 标定过期锁存 === *)
IF (uCalAgeMin >= uCalPeriodMin) AND (uCalPeriodMin > UDINT#0) THEN
    bCalOverdue := TRUE;                          // 到期锁存
    uInfo := 16#0002_06B2;                        // 信息级：过期取样出口闭锁
END_IF
IF _eState = E_DL_AnaPhase.eCal AND bCalDone THEN
    bCalOverdue := FALSE;                         // 标定完成反馈解除锁存（解除路径可达）
END_IF

(* === 段 5 · 主状态机（ENUM + CASE，含 ELSE 兜底）=== *)
CASE _eState OF
E_DL_AnaPhase.eIdle :
    bSampleValid := FALSE;                        // 空闲不出有效
    IF uFault <> 16#0000 THEN
        _eState := E_DL_AnaPhase.eFault;          // 故障优先
    ELSIF bCalReq THEN
        _eState := E_DL_AnaPhase.eCal;            // 标定命令最高优先
    ELSIF bPurgeReqEff THEN
        _eState := E_DL_AnaPhase.ePurge;          // 吹扫次优先
    ELSIF bSampleReqEff AND (NOT bCalOverdue) THEN
        _eState := E_DL_AnaPhase.eSample;         // 取样联锁前置：过期禁取样
    END_IF

E_DL_AnaPhase.eSample :
    bSampleValid := FALSE;                        // 取样中出口未有效（相完成才有效）
    IF uFault <> 16#0000 THEN
        bAbortSample := TRUE;                     // 故障打断取样（仅故障可打断，禁其他相打断）
        _eState := E_DL_AnaPhase.eFault;          // 转故障相
    ELSIF fbSeq.nCurrentStep = 1 THEN
        _eState := E_DL_AnaPhase.ePurge;          // 顺控推到吹扫步：转吹扫相（先完成当前相才切换）
    END_IF

E_DL_AnaPhase.ePurge :
    bSampleValid := FALSE;                        // 吹扫相不出有效
    IF uFault <> 16#0000 THEN
        _eState := E_DL_AnaPhase.eFault;          // 故障转出
    ELSIF bPurgeDone AND bPurgeMinOk THEN
        bSampleValid := TRUE;                     // 吹扫完成且最短时长满足：取样出口有效（本轮吹扫后样本可用）
        _eState := E_DL_AnaPhase.eIdle;           // 回空闲待下轮
    END_IF

E_DL_AnaPhase.eCal :
    bSampleValid := FALSE;                        // 标定相不出有效
    IF uFault <> 16#0000 THEN
        _eState := E_DL_AnaPhase.eFault;          // 故障转出
    ELSIF bCalDone THEN
        bCalOverdue := FALSE;                     // 标定完成解除过期锁存
        _eState := E_DL_AnaPhase.eIdle;           // 回空闲
    END_IF

E_DL_AnaPhase.eFault :
    bSampleValid := FALSE;                        // 故障相闭锁出口
    IF uFault = 16#0000 THEN
        bAbortSample := FALSE;                    // 解锁同步清打断标志
        _eState := E_DL_AnaPhase.eIdle;           // 回空闲
    END_IF

ELSE
    _eState := E_DL_AnaPhase.eFault;              // 非法状态拦截
    uFault := 16#0002_06C2;                       // 故障级：相 ID 越界复用组态码段
END_CASE

(* === 段 6 · 输出映射 === *)
bError := (uFault <> 16#0000);                    // 故障标志仅由故障级码置位（R45 配对）
IF bError THEN
    uErrorId := uFault;                           // 故障级优先上报
ELSE
    uErrorId := uInfo;                            // 否则上报信息级码
END_IF
ePhaseOut := _eState;                             // 输出枚举段尾单点映射（N2 规则）
END_FUNCTION_BLOCK

(* ---- FB_DL_AndonLinePack.st ---- *)
(*
  Component : FB_DL_AndonLinePack
  Category  : DL_Process
  Type      : FB
  Version   : 1.0.0
  CodeSeg   : 16#06_0_40
  Summary   : 包装线安灯分级呼叫与响应报表：三级呼叫仲裁锁存 + 呼叫/应答/解除三段独立计时 + 台账。
              Andon line pack: three-level call arbitration latch, independent call/ack/clear timers, response ledger.
  溯源声明  : 仅借 t2-isa182 安灯呼叫分级与报表口径域，代码 clean-room（T2 借鉴件）
  边界安全  : 三段计时（呼叫→应答→解除）各自独立 TON 实例，禁止共用（按派单要点）；
              仲裁锁存：高级别呼叫可抢占低级别，解除路径可达（对应级别复位指令沿）；
              响应/解除超时为非锁存提示；呼叫/应答计数走沿防电平重复累加；计数防回卷；
              CASE 必带 ELSE 兜底；TON 每拍无条件刷新（段 0）。
  复用      : 复用 FB_DL_AndonCallSystem 仲裁语义 + FB_DL_RuntimeMeter 台账口径（clean-room 自含实现，无实例依赖）
*)

FUNCTION_BLOCK FB_DL_AndonLinePack
VAR_INPUT
    bRun      : BOOL;                   (* 安灯使能 · Enable *)
    bCallL1   : BOOL;                   (* 一级呼叫 [事件]，轻微 · Level 1 call *)
    bCallL2   : BOOL;                   (* 二级呼叫 [事件]，一般 · Level 2 call *)
    bCallL3   : BOOL;                   (* 三级呼叫 [事件]，紧急 · Level 3 call *)
    bAckCmd   : BOOL;                   (* 应答指令 [事件]，沿触发 · Ack command, edge *)
    bClearCmd : BOOL;                   (* 解除指令 [事件]，沿触发 · Clear command, edge *)
    tAckLimMs : TIME  := T#60000MS;     (* 呼叫→应答超时阈 [ms] · Ack timeout limit *)
    tClrLimMs : TIME  := T#300000MS;    (* 应答→解除超时阈 [ms] · Clear timeout limit *)
    fEps      : LREAL := 1.0E-6;        (* 浮点判零容差 [实数域] · Floating zero tolerance *)
END_VAR
VAR_OUTPUT
    eActive : (eAlNone := 0, eAlL1 := 1, eAlL2 := 2, eAlL3 := 3);   (* 激活级别枚举输出 / Active level output enum *)
    bAcked  : BOOL;                     (* 已应答标志 [开关] · Acked flag *)
    bAckTmOut: BOOL;                    (* 呼叫→应答超时提示（非锁存）· Ack timeout hint *)
    bClrTmOut: BOOL;                    (* 应答→解除超时提示（非锁存）· Clear timeout hint *)
    nRespCnt: UDINT;                    (* 超时响应累计 [次]，防回卷 · Timeout response count *)
    nCloseCnt: UDINT;                   (* 正常解除累计 [次]，防回卷 · Normal close count *)
    bError  : BOOL;                     (* 故障标志，与故障码配对 · Fault flag paired with codes *)
    uErrorId: UDINT;                    (* 事件码 16#0000_0040，0 无事件 · Event code *)
END_VAR
VAR
    _eState  : (eStCalm := 0, eStCalling := 1, eStAcked := 2);   (* 内部状态机 / Internal state machine *)
    _nLevel  : INT;     (* 内部激活级别 [级]，与输出枚举分离 / Internal level *)
    uCode    : WORD;    (* 码位暂存，每拍重算 [码] · Code staging *)
    tonAck   : TON;     (* 呼叫→应答计时 [ms]，独立实例 1 · Ack timer, instance 1 *)
    tonClr   : TON;     (* 应答→解除计时 [ms]，独立实例 2 · Clear timer, instance 2 *)
    rTrigAck : R_TRIG;  (* 应答沿检测 · Ack edge *)
    rTrigClr : R_TRIG;  (* 解除沿检测 · Clear edge *)
    bCallNow : BOOL;    (* 仲裁后呼叫有效 [开关] · Arbitrated call active *)
    bAckTmPrv: BOOL;    (* 上拍应答超时提示快照，沿判据 · Previous ack hint snapshot *)
    bClrTmPrv: BOOL;    (* 上拍解除超时提示快照，沿判据 · Previous clear hint snapshot *)
    nCycles  : UDINT;   (* 呼叫周期计数 [次]，防回卷 · Call cycle count *)
END_VAR
VAR CONSTANT
    DL_ALP_WRAP : UDINT := 4294967290;  (* 计数防回卷余量 [次] · Counter wrap guard *)
END_VAR

(* === 段 0 · 实例刷新（每拍无条件，红线 7）=== *)
tonAck(IN := (_eState = eStCalling), PT := tAckLimMs);  (* 呼叫→应答独立计时 / Independent ack timer *)
tonClr(IN := (_eState = eStAcked), PT := tClrLimMs);    (* 应答→解除独立计时 / Independent clear timer *)
rTrigAck(CLK := bAckCmd);                               (* 应答沿检测 / Ack edge *)
rTrigClr(CLK := bClearCmd);                             (* 解除沿检测 / Clear edge *)

(* === 段 1 · 输入校验与量程闸 === *)
uCode := 16#0000;                       // 每拍清码（可达清零基线）/ Clear codes each scan
IF (tAckLimMs <= T#0MS) OR (tClrLimMs <= T#0MS) THEN
    uCode := 16#0040;                   // 故障级：超时阈非正域 / Fault: non-positive timeout limits
END_IF

(* === 段 2 · 主逻辑：三级仲裁与状态机 === *)
(* 仲裁：高级别抢占，同级不重复计数 / Arbitrate: higher level preempts *)
IF bCallL3 THEN
    bCallNow := TRUE;                   (* 三级最高优先 / Level 3 first *)
    IF _nLevel < 3 THEN
        _nLevel := 3;                   (* 抢占升级 / Preempt to level 3 *)
        IF nCycles < DL_ALP_WRAP THEN
            nCycles := nCycles + 1;     (* 新呼叫周期计数 / Count the new call *)
        END_IF
    END_IF
ELSIF bCallL2 THEN
    bCallNow := TRUE;
    IF _nLevel < 2 THEN
        _nLevel := 2;
        IF nCycles < DL_ALP_WRAP THEN
            nCycles := nCycles + 1;
        END_IF
    END_IF
ELSIF bCallL1 THEN
    bCallNow := TRUE;
    IF _nLevel < 1 THEN
        _nLevel := 1;
        IF nCycles < DL_ALP_WRAP THEN
            nCycles := nCycles + 1;
        END_IF
    END_IF
ELSE
    bCallNow := FALSE;                  (* 无呼叫 / No call *)
END_IF
CASE _eState OF
    eStCalm:                            (* 平静相：无激活告警 / Calm: no active alarm *)
        IF bCallNow AND bRun THEN
            _eState := eStCalling;      (* 拍 N 呼叫进入，拍 N+1 呼叫相 / To calling *)
        END_IF
    eStCalling:                         (* 呼叫相：等应答，超时提示非锁存 / Calling: await ack *)
        IF rTrigAck.Q THEN
            _eState := eStAcked;        (* 拍 N 应答沿，拍 N+1 已应答相 / To acked *)
        ELSIF (NOT bCallNow) THEN
            _eState := eStCalm;         (* 呼叫源撤清回平静（可达解除路径 1）/ Call source gone *)
            _nLevel := 0;               (* 级别清零 / Clear the level *)
        ELSIF tonAck.Q THEN
            bAckTmOut := TRUE;          (* 超时提示（非锁存，本拍置位）/ Timeout hint this scan *)
        END_IF
    eStAcked:                           (* 已应答相：等解除 / Acked: await clear *)
        IF rTrigClr.Q THEN
            _eState := eStCalm;         (* 解除回平静（可达解除路径 2）/ Clear to calm *)
            _nLevel := 0;
            IF nCloseCnt < DL_ALP_WRAP THEN
                nCloseCnt := nCloseCnt + 1;     (* 正常解除计数 / Count the normal close *)
            END_IF
        ELSIF tonClr.Q THEN
            bClrTmOut := TRUE;          (* 解除超时提示（非锁存）/ Clear timeout hint *)
        END_IF
ELSE
    _eState := eStCalm;                 (* ELSE 兜底回平静相 / ELSE fallback to calm *)
    _nLevel := 0;
END_CASE

(* === 段 3 · 输出映射与故障码（CASE 内未触碰输出枚举）=== *)
eActive := eAlNone;                     (* 级别映射默认 / Default mapping *)
IF _eState <> eStCalm THEN
    IF _nLevel = 3 THEN
        eActive := eAlL3;               (* 三级映射 / Map level 3 *)
    ELSIF _nLevel = 2 THEN
        eActive := eAlL2;               (* 二级映射 / Map level 2 *)
    ELSIF _nLevel = 1 THEN
        eActive := eAlL1;               (* 一级映射 / Map level 1 *)
    END_IF
END_IF
bAcked := (_eState = eStAcked);         (* 已应答标志 / Acked flag *)
IF (NOT bCallNow) AND (_eState = eStCalm) THEN
    bAckTmOut := FALSE;                 (* 超时提示可达清零 / Reachable clear of hints *)
    bClrTmOut := FALSE;
END_IF
IF NOT bRun THEN
    _eState := eStCalm;                 (* 撤使能回平静（可达解除路径 3）/ Disable to calm *)
    _nLevel := 0;
END_IF
IF bAckTmOut AND (NOT bAckTmPrv) THEN
    IF nRespCnt < DL_ALP_WRAP THEN
        nRespCnt := nRespCnt + 1;       (* 超时响应上升沿计数，防电平重复累加 / Edge-counted timeout responses *)
    END_IF
END_IF
IF bClrTmOut AND (NOT bClrTmPrv) THEN
    IF nRespCnt < DL_ALP_WRAP THEN
        nRespCnt := nRespCnt + 1;       (* 解除超时上升沿计数 / Edge-counted clear timeouts *)
    END_IF
END_IF
bAckTmPrv := bAckTmOut;                 (* 提示快照更新 / Update the hint snapshots *)
bClrTmPrv := bClrTmOut;
bError := (uCode <> 16#0000);           (* 故障标志配对 / Fault flag paired *)
uErrorId := WORD_TO_UDINT(uCode);       (* 码位单点写入（16#0000_0040 形态）/ Single write point *)
END_FUNCTION_BLOCK

(* ---- FB_DL_AndonRespTimeReport.st ---- *)
(*
  FB_DL_AndonRespTimeReport  —  安灯呼叫→应答→解除三段计时与四级响应分档 / Andon call-ack-clear timing with four response buckets
  分类 Category : DL_Process
  码位 Code     : 16#06_0_89
  版本 Version  : 1.0.0
  溯源 Source   : OMAC PackML + ISA-18.2 语义借鉴 · clean-room 实现，仅借分类/参数域/命名，未复制源码
  功能 Function : 1) 呼叫→应答→解除三段各自计时，每段计时器在进入相时复位，防上一轮残值续累；
                  2) 响应时长按四级门限分档，附各档累计计数与应答样本分母；
                  3) 呼叫未应答即解除时不计入应答时长统计（应答样本分母单独计数，口径显式）。
  边界 Boundary : ① 三段计时器各自在进入相时复位（tCallDur / tAckDur / tClearDur 置 0）；
                  ② 未应答即解除不计入应答时长统计（nAckSamples 为分母，显式输出）；
                  ③ 分档边界两条验收向量见下方「验收向量」段（正好整除 / 上限+1）；
                  ④ 结论三行同向：当前段计时 → 分档等级 → 活动标志。
  依赖 Depends  : None

  验收向量（分档边界，TIME 门限 5s / 15s / 30s）:
    V1 正好整除：应答时长 = 5.000 s → 等级 1（取 <= 门限，闭区间）；
    V2 上限 +1  ：应答时长 = 5.001 s → 等级 2；
    V3 上限 +1  ：应答时长 = 30.001 s → 等级 4；
    V4 未应答解除：tCallDur 计入、nAckSamples 不增、tAckDur 保持 0。
  码表 Error codes（本件子码步进 16#10，避让邻件码位）:
    16#0002_0689 故障级：分档门限非严格递增（须 L1 < L2 < L3）
    16#0002_0699 故障级：相 ID 越界（枚举兜底路径）
    16#0002_06A9 信息级：未应答即解除，本次不计入应答时长统计（不置 bError）
*)

TYPE E_DL_AndonPhase :
(
    eIdle     := 0,   // 空闲 / Idle
    eCalling  := 10,  // 呼叫中（等应答）/ Calling, waiting for ack
    eAcked    := 20,  // 已应答（等解除）/ Acknowledged, waiting for clear
    eCleared  := 30,  // 已解除（本轮结束）/ Cleared, round finished
    eFault    := 90   // 故障锁定 / Fault locked
);
END_TYPE

FUNCTION_BLOCK FB_DL_AndonRespTimeReport
VAR_INPUT
    bEnable      : BOOL;                          // 总使能，FALSE 回空闲 / Master enable
    bReset       : BOOL;                          // 复位，上升沿清故障与台账 / Reset, clears fault and ledger
    bCall        : BOOL;                          // 安灯呼叫信号（电平）/ Andon call signal, level
    bAck         : BOOL;                          // 应答信号（电平）/ Acknowledgement signal
    bClear       : BOOL;                          // 呼叫解除信号（电平）/ Call clear signal
    tCycle       : TIME := T#10MS;                // 任务周期 [ms]，计时累加步长 / Task cycle [ms]
    atLvlLimit   : ARRAY[1..3] OF TIME;           // 四级分档门限 [ms]，须严格递增 / Four-level bucket limits [ms]
    tAckTimeout  : TIME := T#120S;                // 应答超时 [ms]，0 = 不监控 / Ack timeout [ms]
END_VAR
VAR_OUTPUT
    tCallDur     : TIME;                          // 本轮呼叫时长 [ms]（含未应答轮）/ Current call duration [ms]
    tAckDur      : TIME;                          // 本轮应答时长 [ms] / Current response duration [ms]
    tClearDur    : TIME;                          // 本轮解除时长 [ms] / Current clear duration [ms]
    tRespAvg     : TIME;                          // 应答时长累计 [ms]（分母见 nAckSamples）/ Response time total [ms]
    nAckSamples  : INT;                           // 应答样本数 [次]（统计分母，显式）/ Acked sample count, explicit denominator
    nLevel       : INT;                           // 本轮响应分档 1~4，0 = 无结论 / Response bucket 1..4, 0 = none
    anLvlCount   : ARRAY[1..4] OF INT;            // 各档累计次数 [次] / Per-level counters
    bActive      : BOOL;                          // 呼叫活动标志 / Call active flag
    bAckTimeout  : BOOL;                          // 应答超时标志（保持型）/ Ack timeout, held
    bError       : BOOL;                          // 故障标志，与故障级码配对 / Fault flag paired with fault codes
    uErrorId     : UDINT;                         // 事件码，0 = 无事件 / Event code, 0 = none
    eStateOut    : E_DL_AndonPhase;               // 状态机当前态，段尾单点映射 / Phase mapped at tail
END_VAR
VAR
    _eState      : E_DL_AndonPhase := E_DL_AndonPhase.eIdle;  // 内部状态 / Internal state
    rtrReset     : R_TRIG;                        // 复位沿 / Reset edge
    tonAckTo     : TON;                           // 应答超时计时（无条件刷新）/ Ack timeout timer
    bCfgOk       : BOOL;                          // 门限组态合法 / Bucket limits valid
    bAckCounted  : BOOL;                          // 本轮已计应答样本 / Ack counted this round
    nI           : INT;                           // 台账循环下标 / Ledger loop index
    nLvlBuf      : INT;                           // 分档暂存 / Bucket buffer
    uFault       : UDINT;                         // 锁存故障码 / Latched fault code
    uInfo        : UDINT;                         // 信息级码 / Information code
END_VAR
VAR CONSTANT
    DL_AND_LVLMAX : INT := 4;                     // 分档总数 [档] / Bucket count
    DL_AND_CNTMAX : INT := 32000;                 // 台账计数上限 [次]，防 INT 溢出 / Ledger counter ceiling
END_VAR

(* === 段 0 · 实例刷新（无条件周期调用）=== *)
rtrReset(CLK := bReset);                          // 每拍刷新复位沿
tonAckTo(IN := (_eState = E_DL_AndonPhase.eCalling), PT := tAckTimeout);   // 应答超时计时，无条件刷新

(* === 段 1 · 组态闸：分档门限严格递增 === *)
bCfgOk := (atLvlLimit[1] > T#0MS) AND (atLvlLimit[2] > atLvlLimit[1])
          AND (atLvlLimit[3] > atLvlLimit[2]);   // 严格递增，倒置即组态报码
IF NOT bCfgOk THEN
    uFault := 16#0002_0689;                       // 故障级：分档门限非法
END_IF
IF rtrReset.Q THEN
    uFault := 16#0000;                            // 复位沿清锁存
    bAckTimeout := FALSE;                         // 超时标志同步复位
    FOR nI := 1 TO DL_AND_LVLMAX DO
        anLvlCount[nI] := 0;                      // 台账清零（复位口径显式）
    END_FOR
    nAckSamples := 0;                             // 应答样本分母清零
    tRespAvg := T#0MS;                            // 应答累计清零
END_IF

(* === 段 2 · 主状态机（ENUM + CASE，含 ELSE 兜底）=== *)
CASE _eState OF
E_DL_AndonPhase.eIdle :
    bActive := FALSE;                             // 空闲无活动呼叫
    nLevel := 0;                                  // 分档无结论
    tCallDur := T#0MS;                            // 呼叫计时复位（进入新轮前清零）
    tAckDur := T#0MS;                             // 应答计时复位
    tClearDur := T#0MS;                           // 解除计时复位
    bAckCounted := FALSE;                         // 本轮未计样本
    uInfo := 16#0000;                             // 信息码清零
    IF uFault <> 16#0000 THEN
        _eState := E_DL_AndonPhase.eFault;        // 故障优先
    ELSIF bEnable AND bCall THEN
        tCallDur := T#0MS;                        // 进入呼叫相：计时器复位（防残值续累）
        bActive := TRUE;                          // 活动标志置位
        _eState := E_DL_AndonPhase.eCalling;
    END_IF

E_DL_AndonPhase.eCalling :
    bActive := TRUE;                              // 呼叫活动
    tCallDur := tCallDur + tCycle;                // 呼叫时长累加
    IF bAck THEN
        tCallDur := tCallDur;                     // 呼叫时长定格（本拍不再累加）
        tAckDur := T#0MS;                         // 进入应答相：应答计时器复位
        _eState := E_DL_AndonPhase.eAcked;        // 本拍行为：转已应答相
    ELSIF tonAckTo.Q THEN
        bAckTimeout := TRUE;                      // 置位型：应答超时（段尾不清零）
    ELSIF NOT bCall THEN
        uInfo := 16#0002_06A9;                    // 信息级：未应答即解除，不计入应答统计
        _eState := E_DL_AndonPhase.eCleared;      // 直接转解除相（分母口径不污染）
    END_IF

E_DL_AndonPhase.eAcked :
    bActive := TRUE;                              // 仍在处理中
    tAckDur := tAckDur + tCycle;                  // 应答时长累加
    IF NOT bAckCounted THEN
        tRespAvg := tRespAvg + tAckDur;           // 应答时长累计入台账
        nAckSamples := nAckSamples + 1;           // 分母 +1（显式口径）
        bAckCounted := TRUE;                      // 本轮已计样本，防重复累加
    END_IF
    IF (NOT bCall) OR bClear THEN
        tClearDur := T#0MS;                       // 进入解除相：解除计时器复位
        _eState := E_DL_AndonPhase.eCleared;      // 转解除相
    END_IF

E_DL_AndonPhase.eCleared :
    tClearDur := tClearDur + tCycle;              // 解除时长累加
    IF NOT bCall THEN
        bActive := FALSE;                         // 呼叫已撤销：活动标志落 0（三行同向）
        IF tAckDur <= atLvlLimit[1] THEN
            nLvlBuf := 1;                         // 分档 1：应答 <= L1（闭区间，正好整除落在本级）
        ELSIF tAckDur <= atLvlLimit[2] THEN
            nLvlBuf := 2;                         // 分档 2：L1 < 应答 <= L2
        ELSIF tAckDur <= atLvlLimit[3] THEN
            nLvlBuf := 3;                         // 分档 3：L2 < 应答 <= L3
        ELSE
            nLvlBuf := DL_AND_LVLMAX;             // 分档 4：应答 > L3（上限 +1 落最高档）
        END_IF
        nLevel := nLvlBuf;                        // 分档结果输出
        IF (nLvlBuf >= 1) AND (nLvlBuf <= DL_AND_LVLMAX) THEN
            IF anLvlCount[nLvlBuf] < DL_AND_CNTMAX THEN
                anLvlCount[nLvlBuf] := anLvlCount[nLvlBuf] + 1;   // 台账计数，饱和防溢出
            END_IF
        END_IF
        _eState := E_DL_AndonPhase.eIdle;         // 本轮结束回空闲（下轮计时器在空闲相复位）
    END_IF

E_DL_AndonPhase.eFault :
    bActive := FALSE;                             // 故障态无活动
    nLevel := 0;                                  // 分档无结论
    IF uFault = 16#0000 THEN
        _eState := E_DL_AndonPhase.eIdle;         // 解锁回空闲
    END_IF

ELSE
    _eState := E_DL_AndonPhase.eFault;            // 非法状态拦截
    uFault := 16#0002_0699;                       // 故障级：相 ID 越界（枚举兜底路径）
    nLevel := 0;                                  // 安全侧无分档
END_CASE
IF NOT bEnable THEN
    _eState := E_DL_AndonPhase.eIdle;             // 失能最高优先回空闲
    bActive := FALSE;                             // 活动标志落 0
    nLevel := 0;                                  // 分档无结论
END_IF

(* === 段 3 · 输出映射（三行同向：段计时 → 分档 → 活动标志）=== *)
IF bCall AND (NOT bActive) THEN
    bActive := TRUE;                              // 呼叫电平与活动标志对齐（防状态机滞后一拍漏报）
END_IF
IF NOT bCall AND (_eState <> E_DL_AndonPhase.eCleared) THEN
    bActive := FALSE;                             // 呼叫撤销且不在解除相：活动标志落 0
END_IF
bError := (uFault <> 16#0000);                    // 故障标志仅由故障级码置位（R45 配对）
IF bError THEN
    uErrorId := uFault;                           // 故障级优先上报
ELSE
    uErrorId := uInfo;                            // 否则上报信息级码
END_IF
eStateOut := _eState;                             // 输出枚举段尾单点映射（N2 规则）
END_FUNCTION_BLOCK
